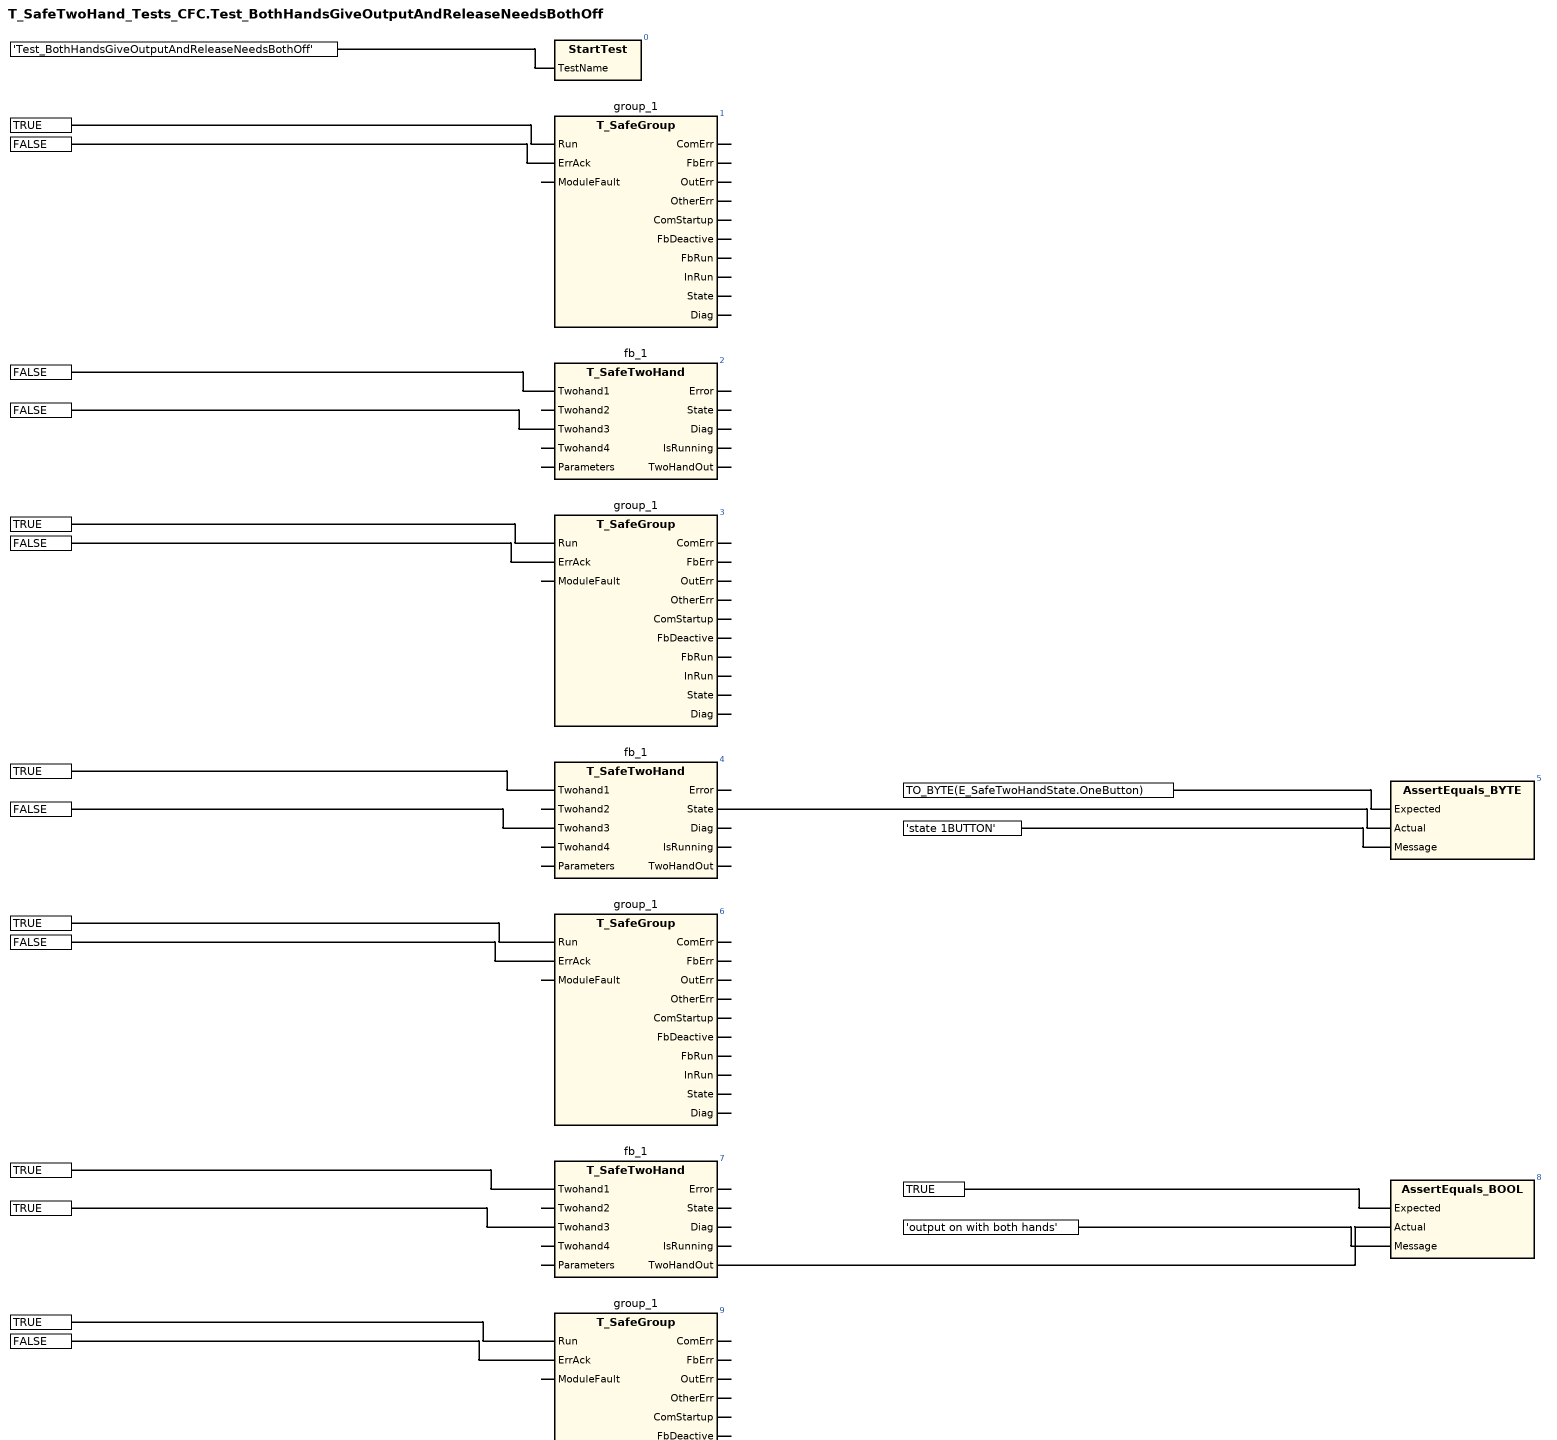
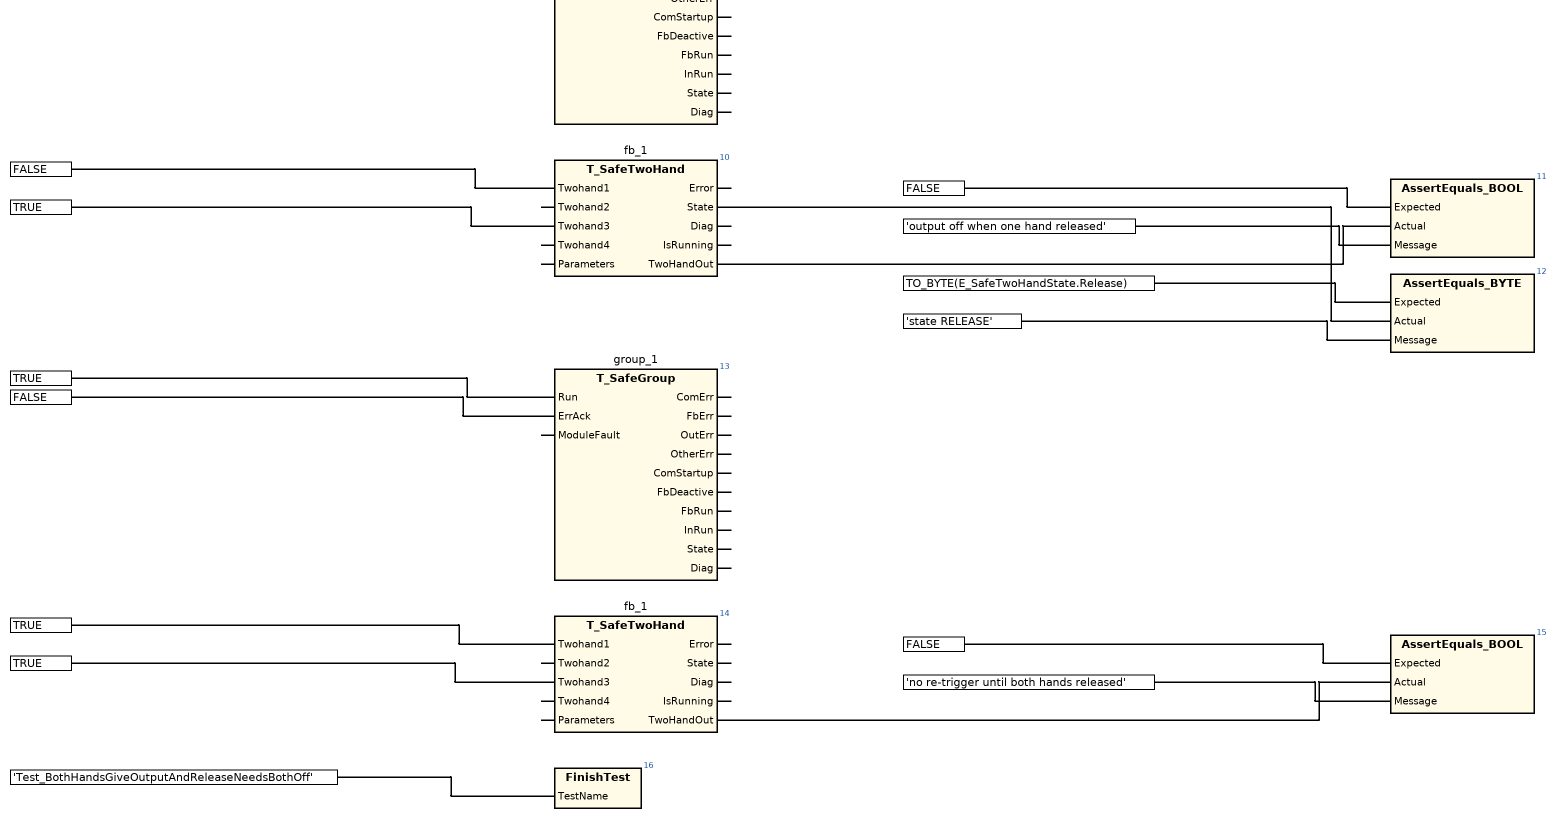
StartTest(TestName := 'Test_BothHandsGiveOutputAndReleaseNeedsBothOff');
group_1(Run := TRUE, ErrAck := FALSE); // T_SafeGroup
fb_1(Twohand1 := FALSE, Twohand3 := FALSE); // T_SafeTwoHand
group_1(Run := TRUE, ErrAck := FALSE); // T_SafeGroup
fb_1(Twohand1 := TRUE, Twohand3 := FALSE); // T_SafeTwoHand
AssertEquals_BYTE(Expected := TO_BYTE(E_SafeTwoHandState.OneButton), Actual := fb_1.State, Message := 'state 1BUTTON');
group_1(Run := TRUE, ErrAck := FALSE); // T_SafeGroup
fb_1(Twohand1 := TRUE, Twohand3 := TRUE); // T_SafeTwoHand
AssertEquals_BOOL(Expected := TRUE, Actual := fb_1.TwoHandOut, Message := 'output on with both hands');
group_1(Run := TRUE, ErrAck := FALSE); // T_SafeGroup
fb_1(Twohand1 := FALSE, Twohand3 := TRUE); // T_SafeTwoHand
AssertEquals_BOOL(Expected := FALSE, Actual := fb_1.TwoHandOut, Message := 'output off when one hand released');
AssertEquals_BYTE(Expected := TO_BYTE(E_SafeTwoHandState.Release), Actual := fb_1.State, Message := 'state RELEASE');
group_1(Run := TRUE, ErrAck := FALSE); // T_SafeGroup
fb_1(Twohand1 := TRUE, Twohand3 := TRUE); // T_SafeTwoHand
AssertEquals_BOOL(Expected := FALSE, Actual := fb_1.TwoHandOut, Message := 'no re-trigger until both hands released');
FinishTest(TestName := 'Test_BothHandsGiveOutputAndReleaseNeedsBothOff');
END_METHOD

METHOD PRIVATE Test_HandDiscrepancyTimeout
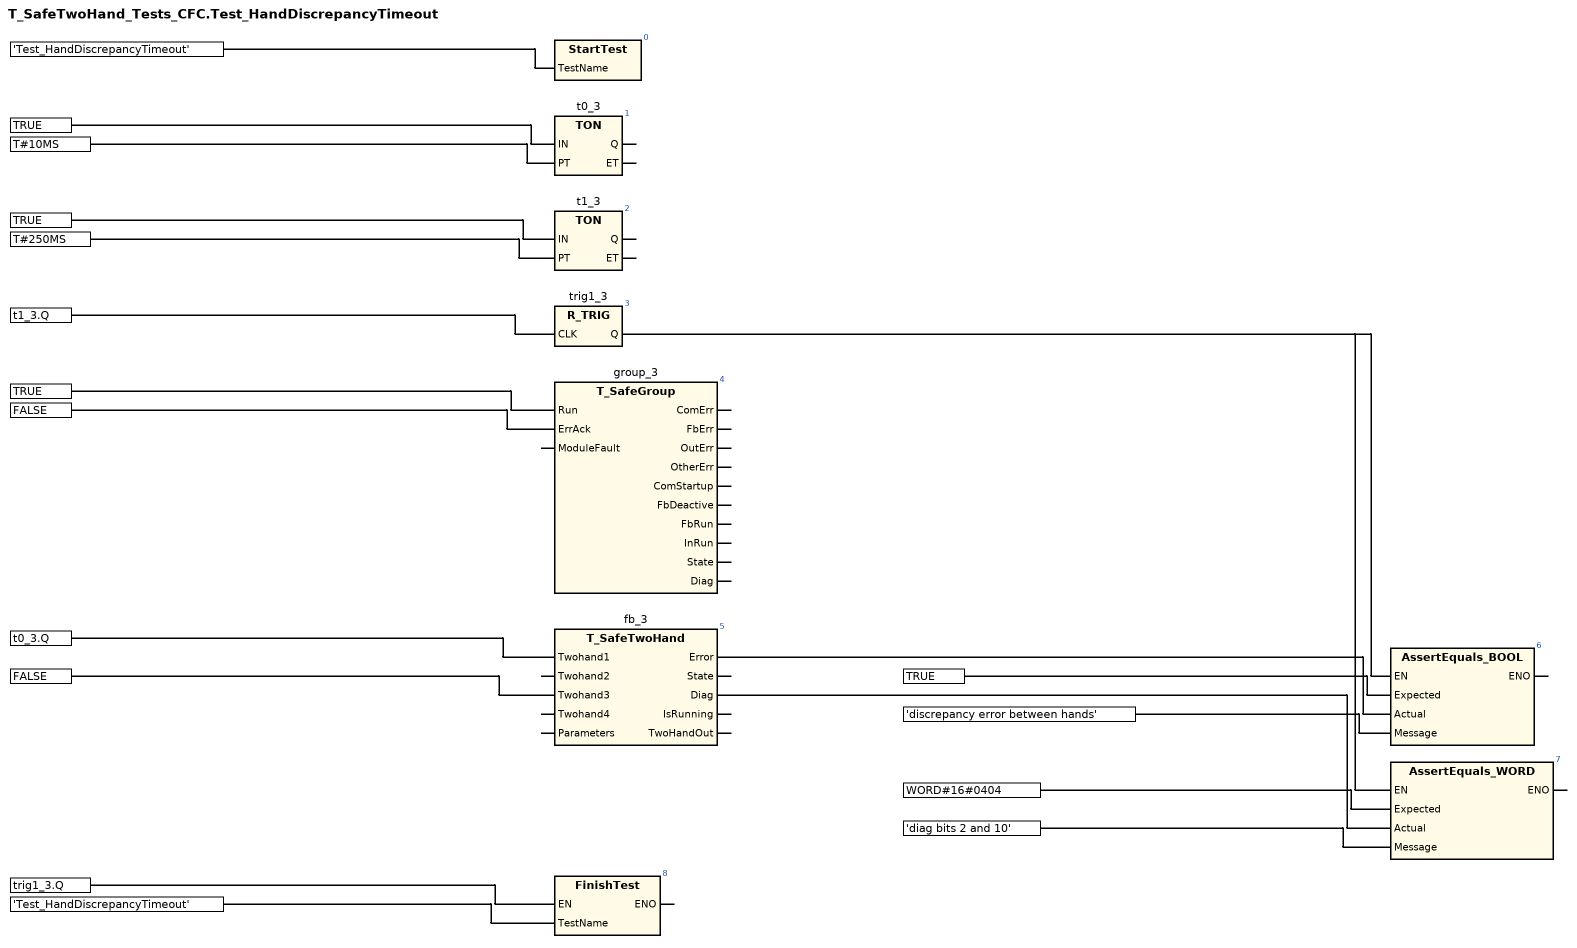
StartTest(TestName := 'Test_HandDiscrepancyTimeout');
t0_3(IN := TRUE, PT := T#10MS); // TON
t1_3(IN := TRUE, PT := T#250MS); // TON
trig1_3(CLK := t1_3.Q); // R_TRIG
group_3(Run := TRUE, ErrAck := FALSE); // T_SafeGroup
fb_3(Twohand1 := t0_3.Q, Twohand3 := FALSE); // T_SafeTwoHand
IF trig1_3.Q THEN AssertEquals_BOOL(Expected := TRUE, Actual := fb_3.Error, Message := 'discrepancy error between hands'); END_IF
IF trig1_3.Q THEN AssertEquals_WORD(Expected := WORD#16#0404, Actual := fb_3.Diag, Message := 'diag bits 2 and 10'); END_IF
IF trig1_3.Q THEN FinishTest(TestName := 'Test_HandDiscrepancyTimeout'); END_IF
END_METHOD

METHOD PRIVATE Test_SecondHandWithoutFirstGivesTwoHandError
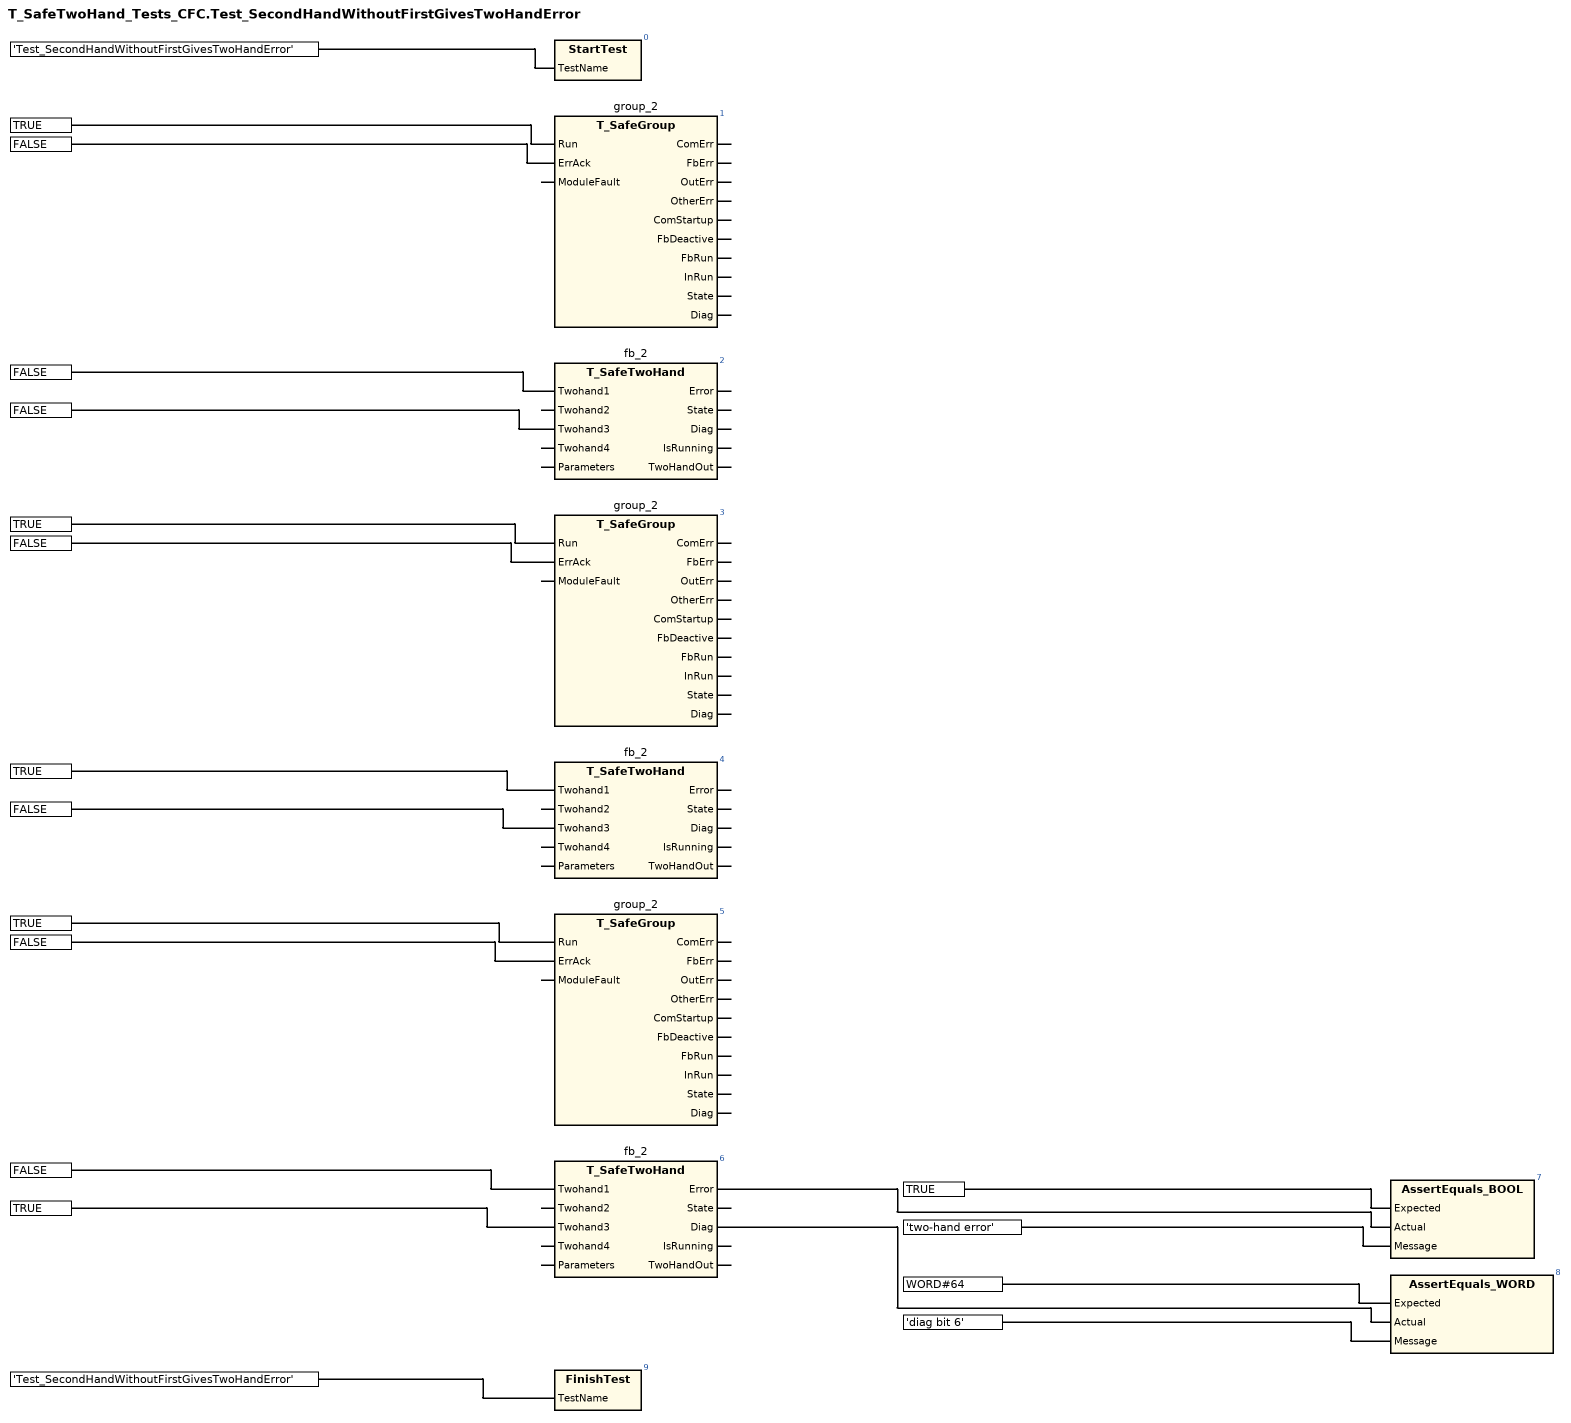
StartTest(TestName := 'Test_SecondHandWithoutFirstGivesTwoHandError');
group_2(Run := TRUE, ErrAck := FALSE); // T_SafeGroup
fb_2(Twohand1 := FALSE, Twohand3 := FALSE); // T_SafeTwoHand
group_2(Run := TRUE, ErrAck := FALSE); // T_SafeGroup
fb_2(Twohand1 := TRUE, Twohand3 := FALSE); // T_SafeTwoHand
group_2(Run := TRUE, ErrAck := FALSE); // T_SafeGroup
fb_2(Twohand1 := FALSE, Twohand3 := TRUE); // T_SafeTwoHand
AssertEquals_BOOL(Expected := TRUE, Actual := fb_2.Error, Message := 'two-hand error');
AssertEquals_WORD(Expected := WORD#64, Actual := fb_2.Diag, Message := 'diag bit 6');
FinishTest(TestName := 'Test_SecondHandWithoutFirstGivesTwoHandError');
END_METHOD

END_FUNCTION_BLOCK

// Tests/T_SafeMuting_Tests_CFC
    // CFC twin of T_SafeMuting_Tests: the same tests drawn as CFC diagrams, the way a TwinSAFE project is authored.
    FUNCTION_BLOCK T_SafeMuting_Tests_CFC EXTENDS T_SafeCfcTestSuite
    VAR
    // Test_OssdBlockedWithoutMutingGivesSafe
    group_1 : T_SafeGroup;
    fb_1 : T_SafeMuting(group := group_1);
    // Test_SequentialMutingKeepsOutputOn
    group_2 : T_SafeGroup;
    fb_2 : T_SafeMuting(group := group_2) := (Parameters := (SequentialInputs := TRUE));
    // Test_SequenceViolationGivesError
    group_3 : T_SafeGroup;
    fb_3 : T_SafeMuting(group := group_3) := (Parameters := (SequentialInputs := TRUE));
    // Test_TwoSensorParallelSequence
    group_4 : T_SafeGroup;
    fb_4 : T_SafeMuting(group := group_4);
END_VAR

Test_OssdBlockedWithoutMutingGivesSafe();
Test_SequentialMutingKeepsOutputOn();
Test_SequenceViolationGivesError();
Test_TwoSensorParallelSequence();

METHOD PRIVATE Test_OssdBlockedWithoutMutingGivesSafe
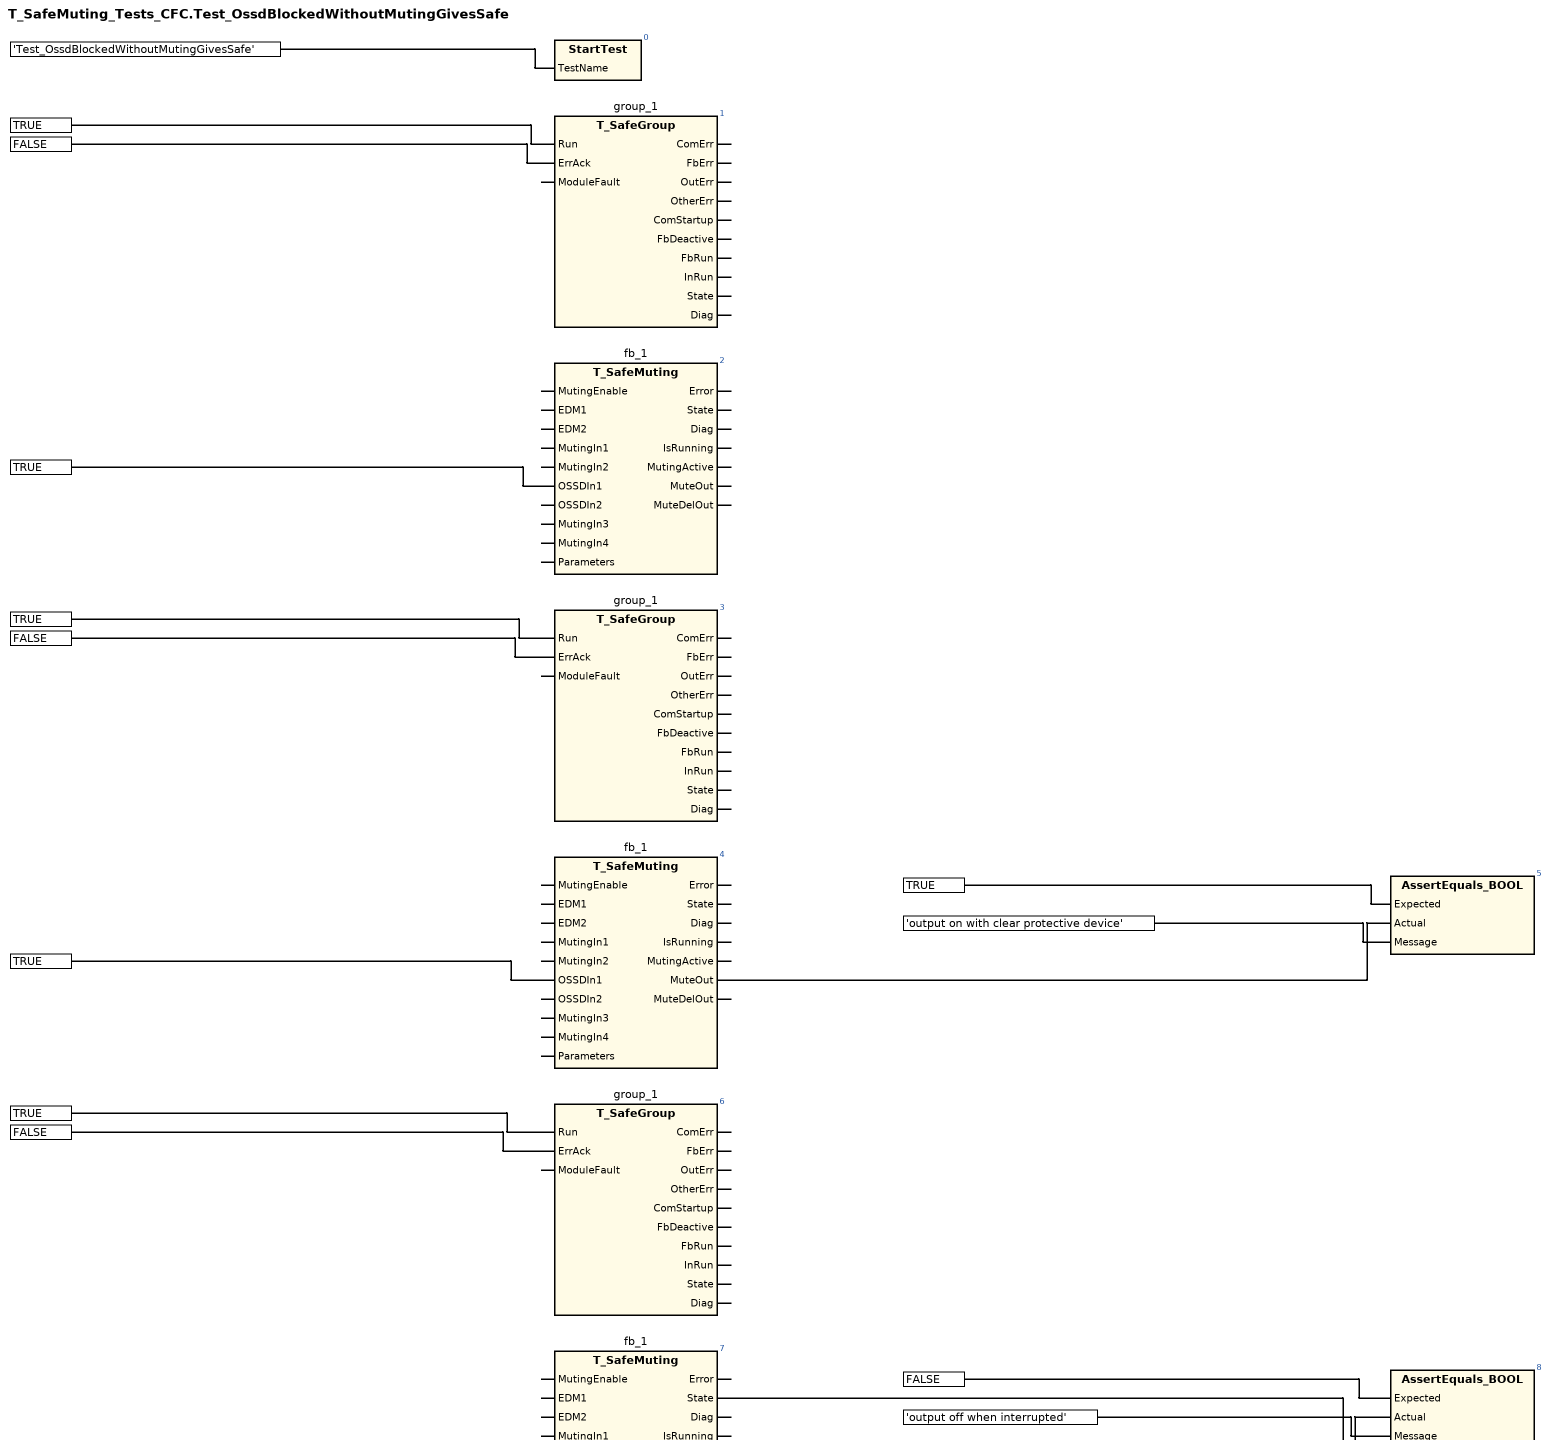
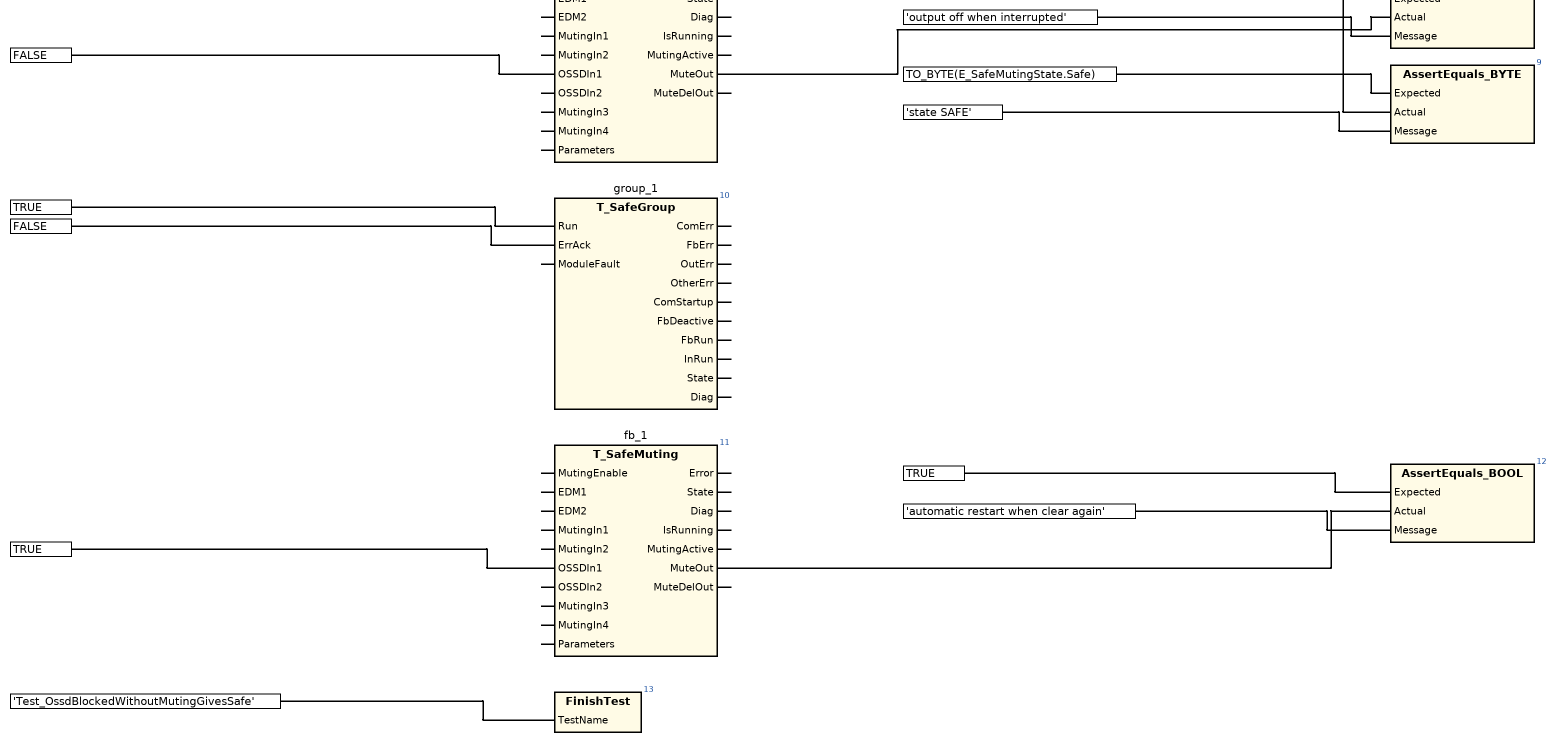
StartTest(TestName := 'Test_OssdBlockedWithoutMutingGivesSafe');
group_1(Run := TRUE, ErrAck := FALSE); // T_SafeGroup
fb_1(OSSDIn1 := TRUE); // T_SafeMuting
group_1(Run := TRUE, ErrAck := FALSE); // T_SafeGroup
fb_1(OSSDIn1 := TRUE); // T_SafeMuting
AssertEquals_BOOL(Expected := TRUE, Actual := fb_1.MuteOut, Message := 'output on with clear protective device');
group_1(Run := TRUE, ErrAck := FALSE); // T_SafeGroup
fb_1(OSSDIn1 := FALSE); // T_SafeMuting
AssertEquals_BOOL(Expected := FALSE, Actual := fb_1.MuteOut, Message := 'output off when interrupted');
AssertEquals_BYTE(Expected := TO_BYTE(E_SafeMutingState.Safe), Actual := fb_1.State, Message := 'state SAFE');
group_1(Run := TRUE, ErrAck := FALSE); // T_SafeGroup
fb_1(OSSDIn1 := TRUE); // T_SafeMuting
AssertEquals_BOOL(Expected := TRUE, Actual := fb_1.MuteOut, Message := 'automatic restart when clear again');
FinishTest(TestName := 'Test_OssdBlockedWithoutMutingGivesSafe');
END_METHOD

METHOD PRIVATE Test_SequenceViolationGivesError
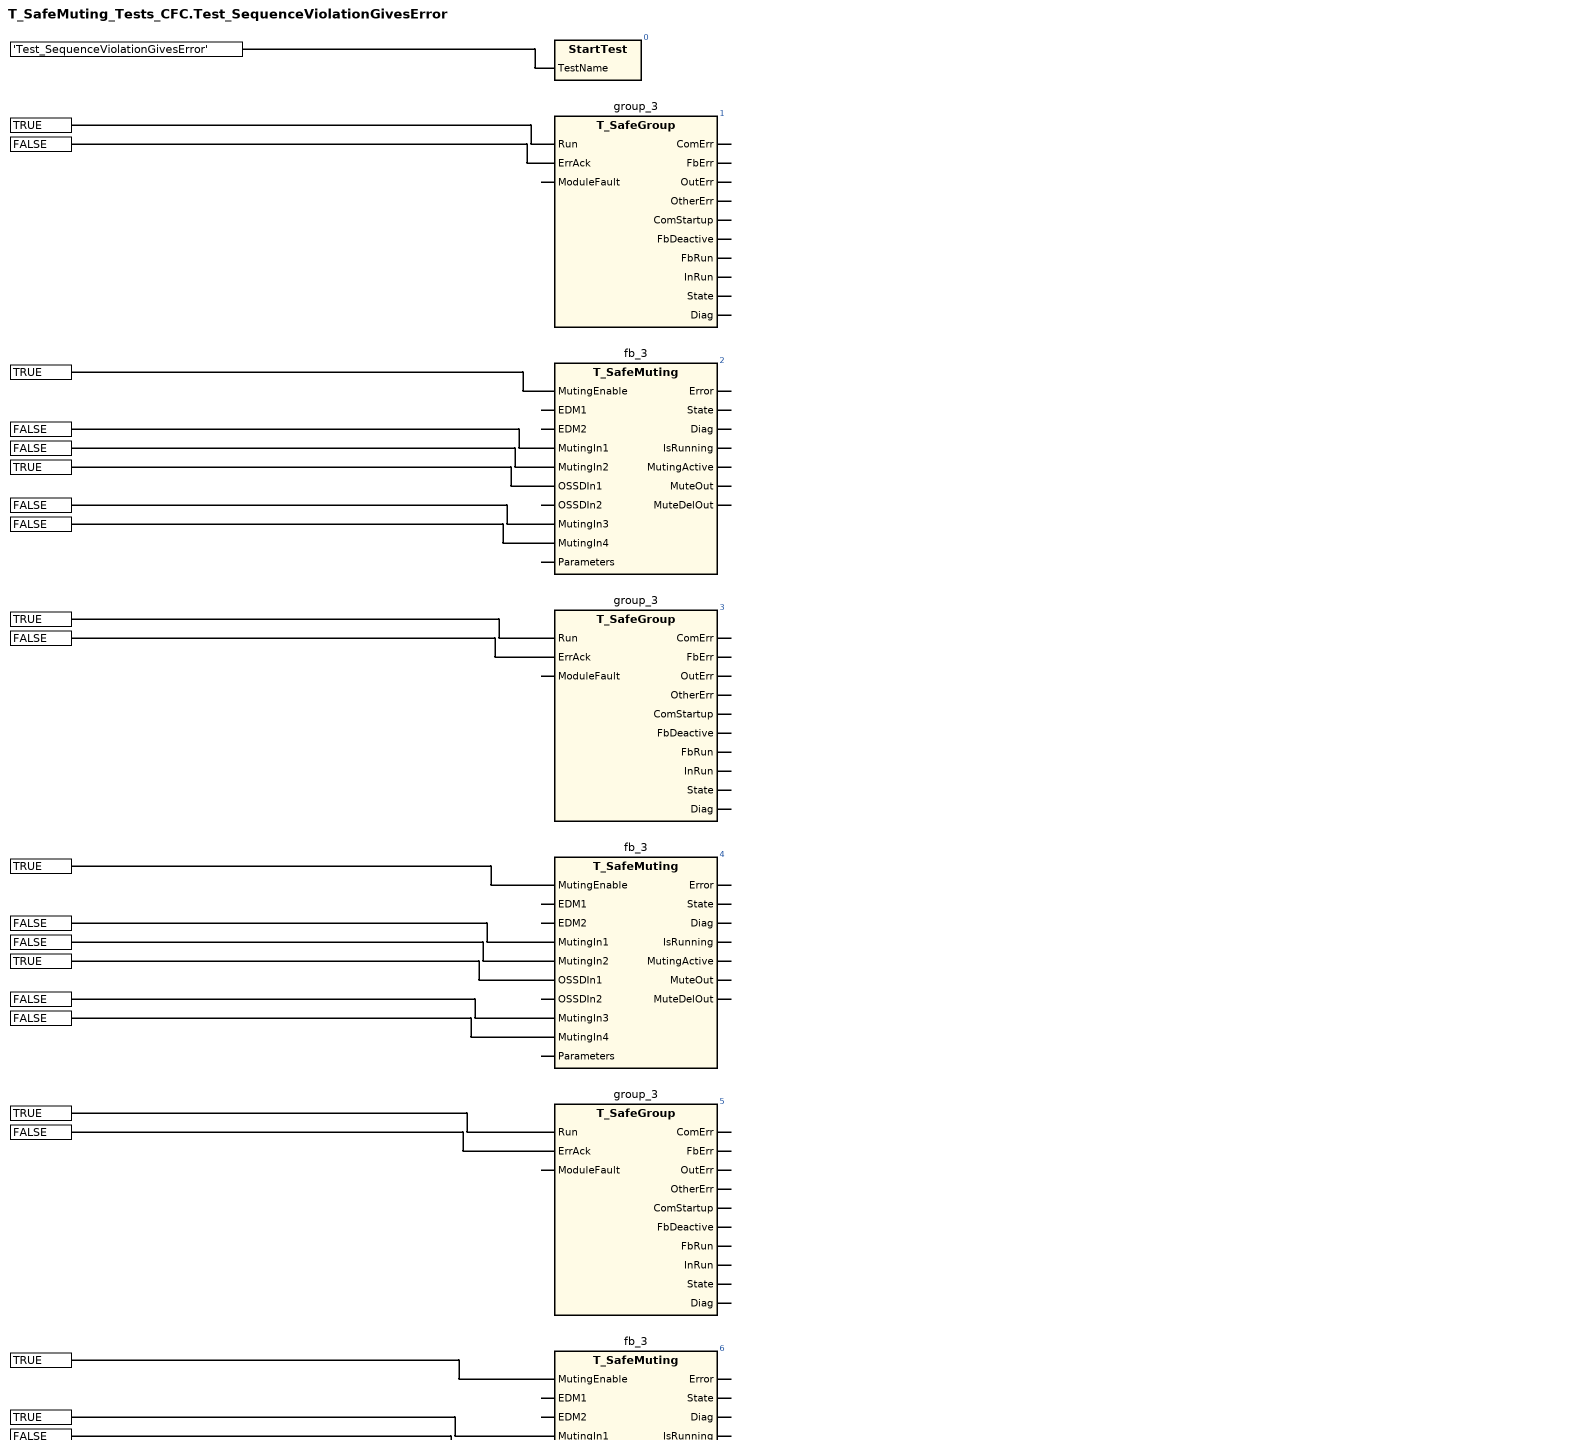
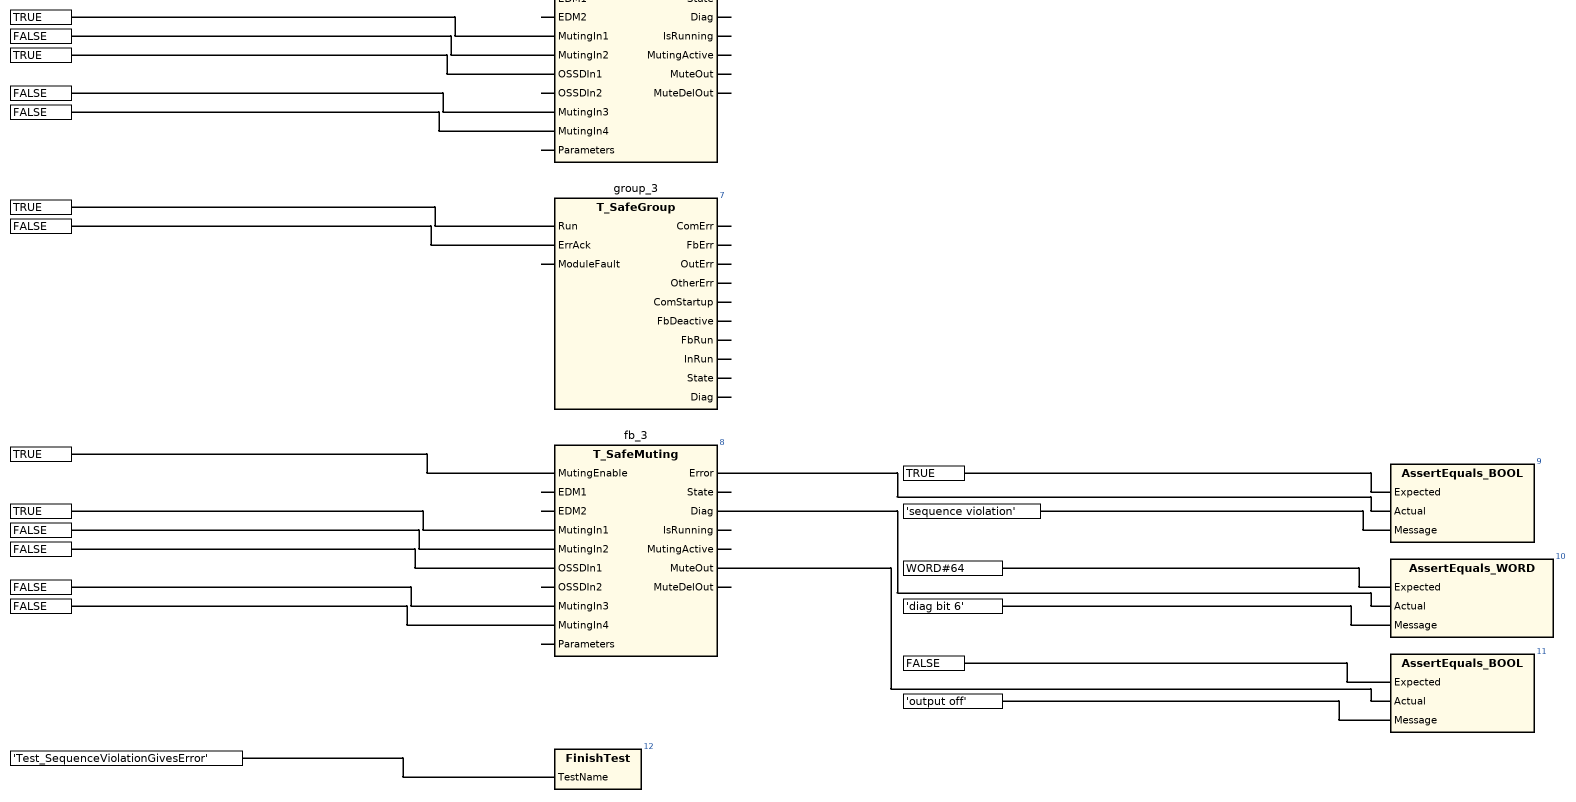
StartTest(TestName := 'Test_SequenceViolationGivesError');
group_3(Run := TRUE, ErrAck := FALSE); // T_SafeGroup
fb_3(
    MutingEnable := TRUE,
    MutingIn1 := FALSE,
    MutingIn2 := FALSE,
    OSSDIn1 := TRUE,
    MutingIn3 := FALSE,
    MutingIn4 := FALSE); // T_SafeMuting
group_3(Run := TRUE, ErrAck := FALSE); // T_SafeGroup
fb_3(
    MutingEnable := TRUE,
    MutingIn1 := FALSE,
    MutingIn2 := FALSE,
    OSSDIn1 := TRUE,
    MutingIn3 := FALSE,
    MutingIn4 := FALSE); // T_SafeMuting
group_3(Run := TRUE, ErrAck := FALSE); // T_SafeGroup
fb_3(
    MutingEnable := TRUE,
    MutingIn1 := TRUE,
    MutingIn2 := FALSE,
    OSSDIn1 := TRUE,
    MutingIn3 := FALSE,
    MutingIn4 := FALSE); // T_SafeMuting
group_3(Run := TRUE, ErrAck := FALSE); // T_SafeGroup
fb_3(
    MutingEnable := TRUE,
    MutingIn1 := TRUE,
    MutingIn2 := FALSE,
    OSSDIn1 := FALSE,
    MutingIn3 := FALSE,
    MutingIn4 := FALSE); // T_SafeMuting
AssertEquals_BOOL(Expected := TRUE, Actual := fb_3.Error, Message := 'sequence violation');
AssertEquals_WORD(Expected := WORD#64, Actual := fb_3.Diag, Message := 'diag bit 6');
AssertEquals_BOOL(Expected := FALSE, Actual := fb_3.MuteOut, Message := 'output off');
FinishTest(TestName := 'Test_SequenceViolationGivesError');
END_METHOD

METHOD PRIVATE Test_SequentialMutingKeepsOutputOn
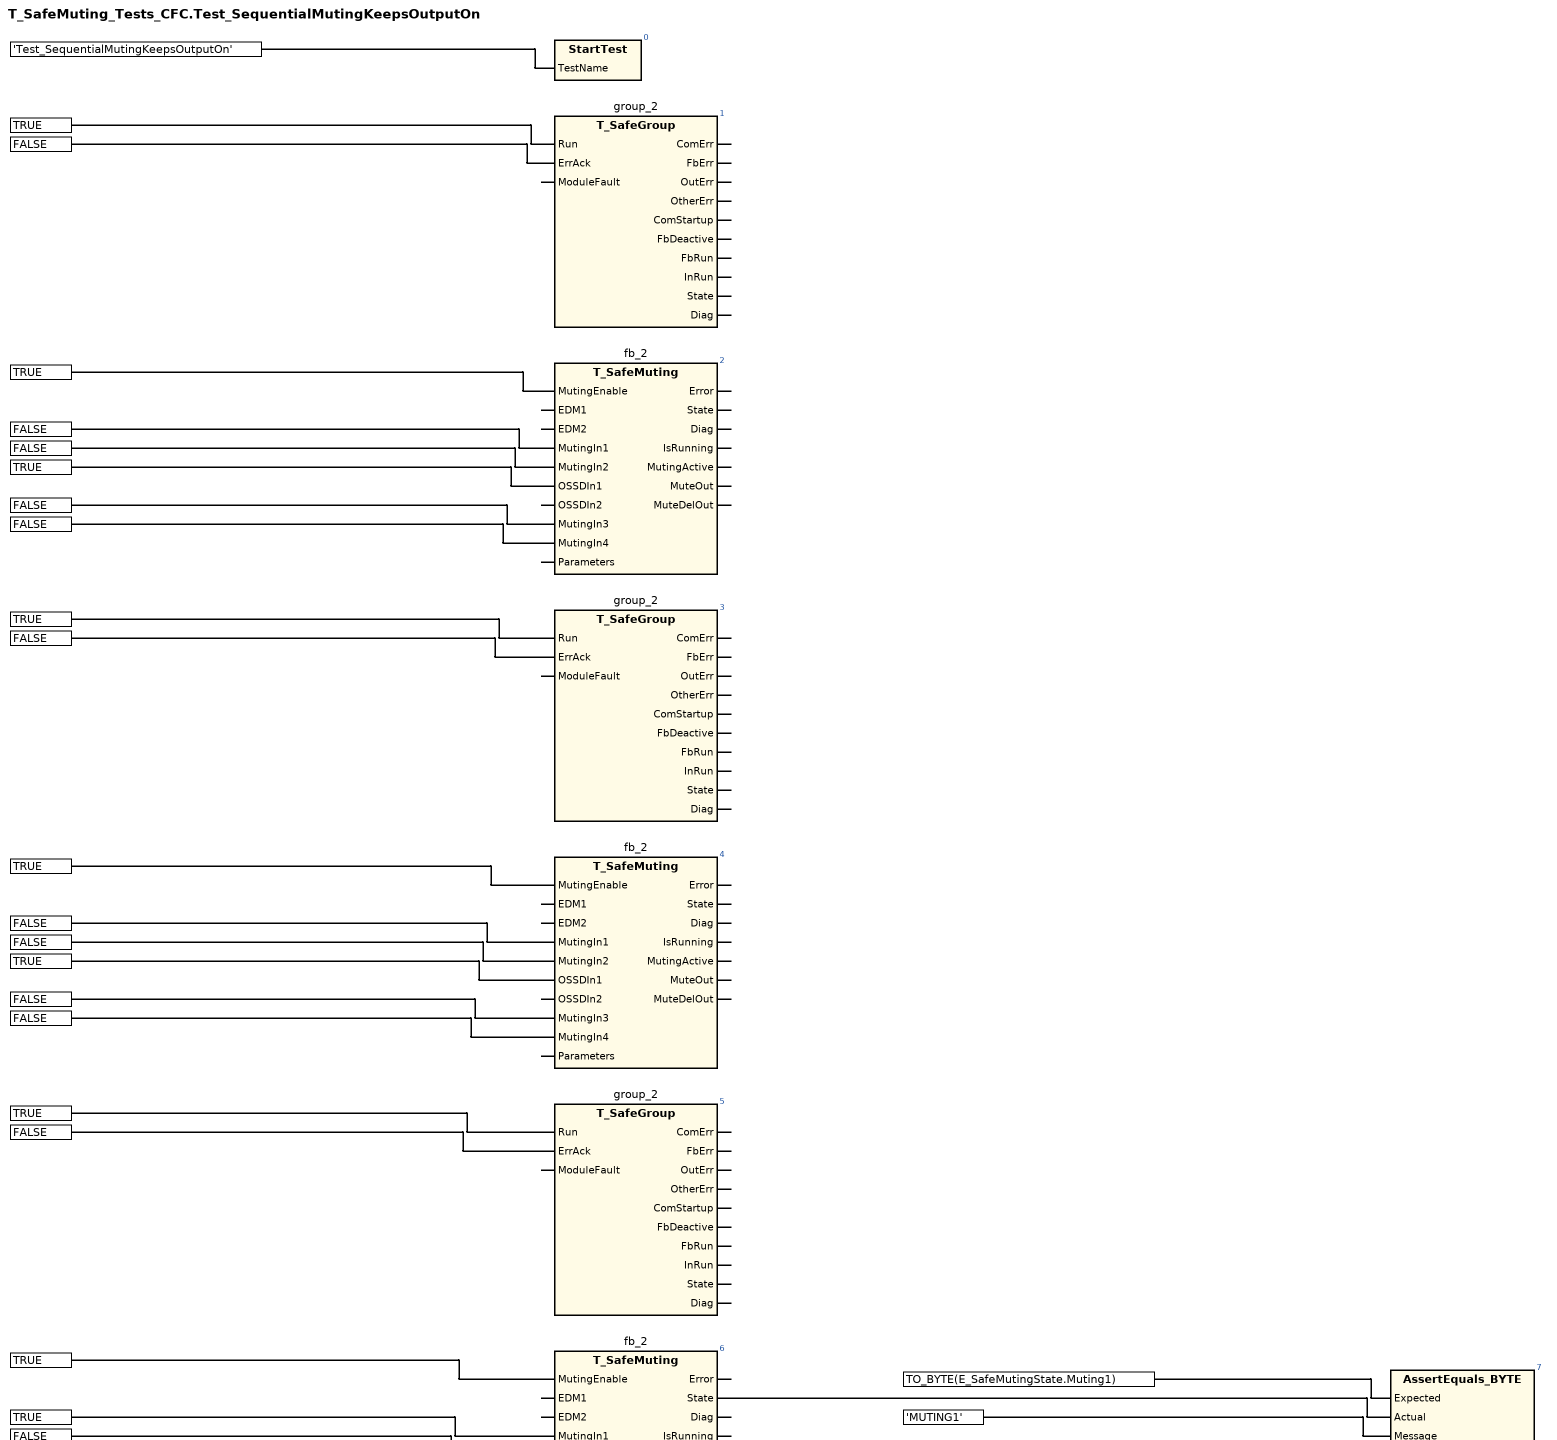
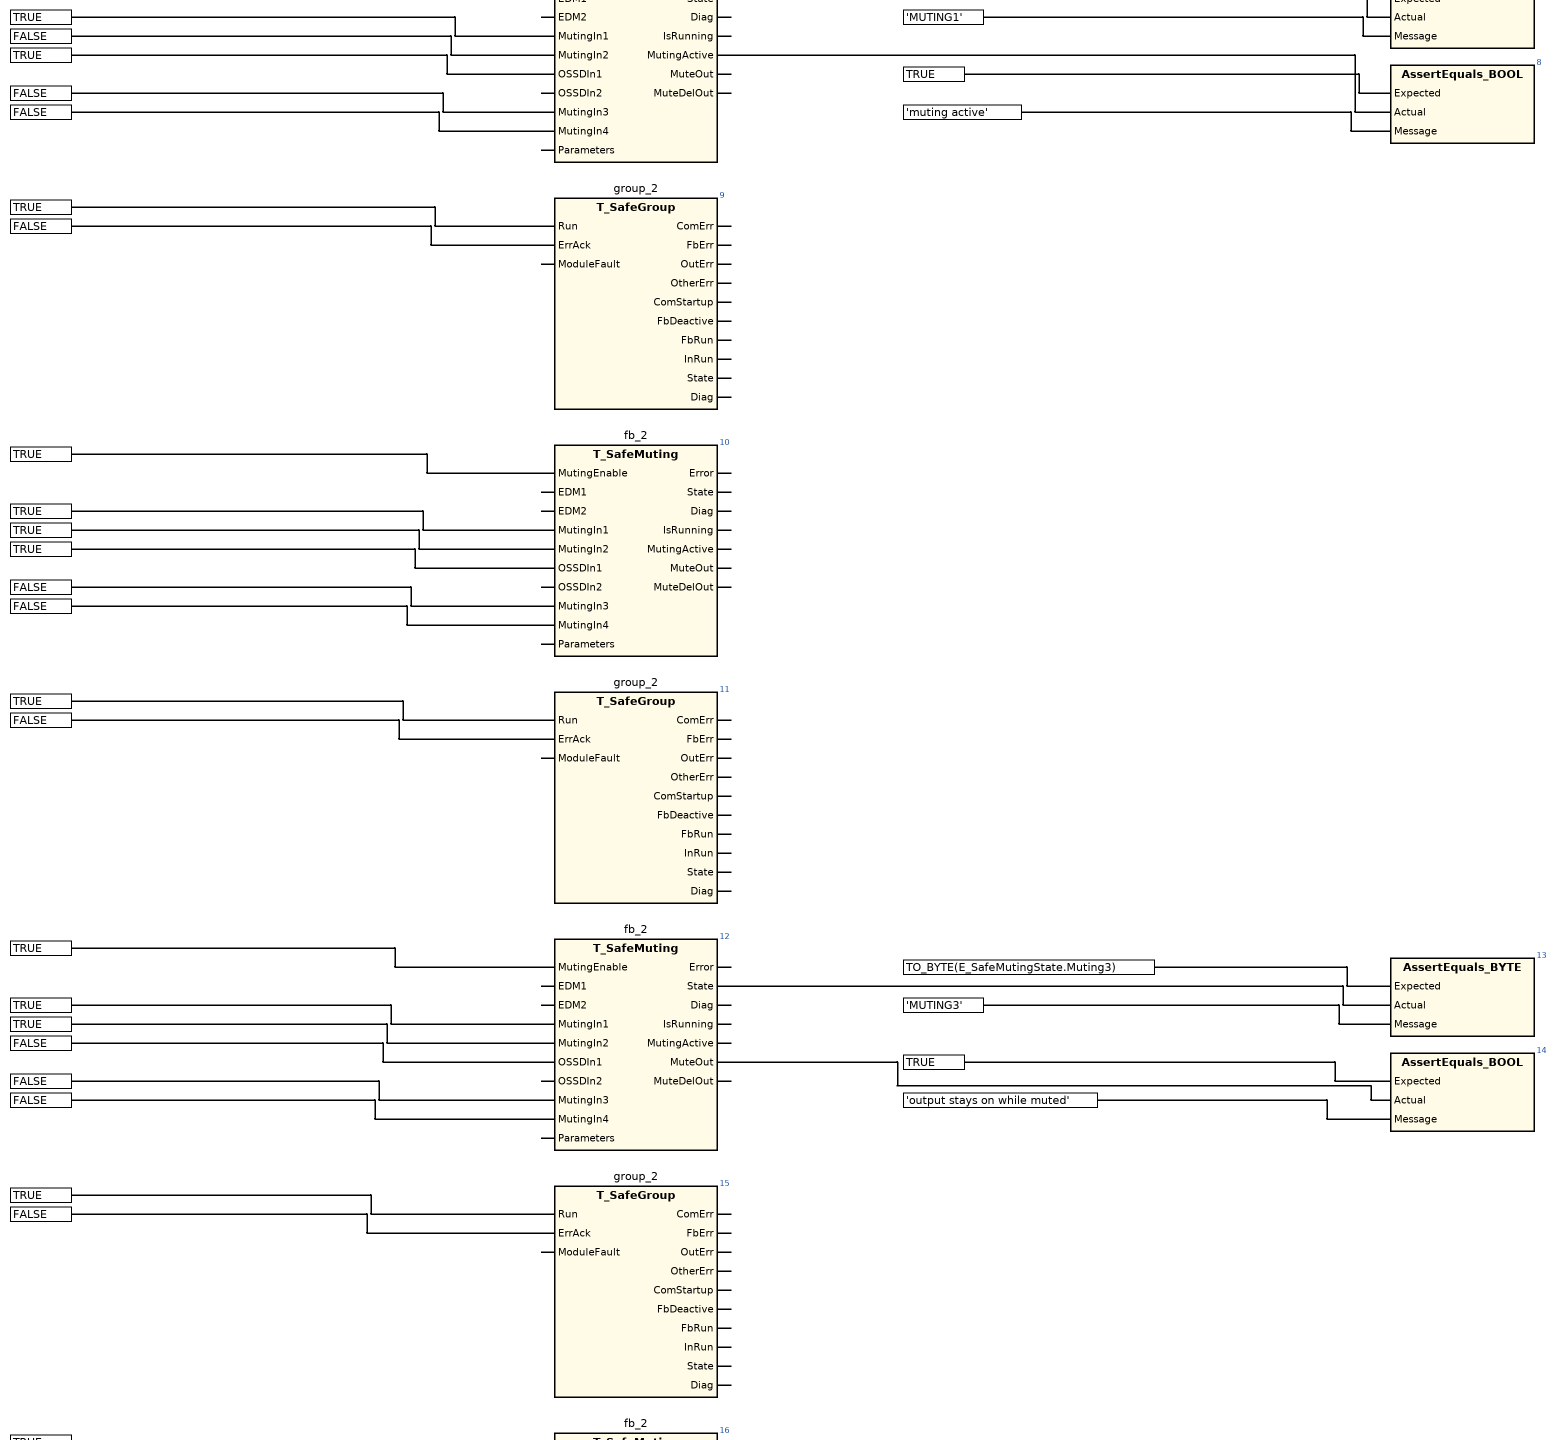
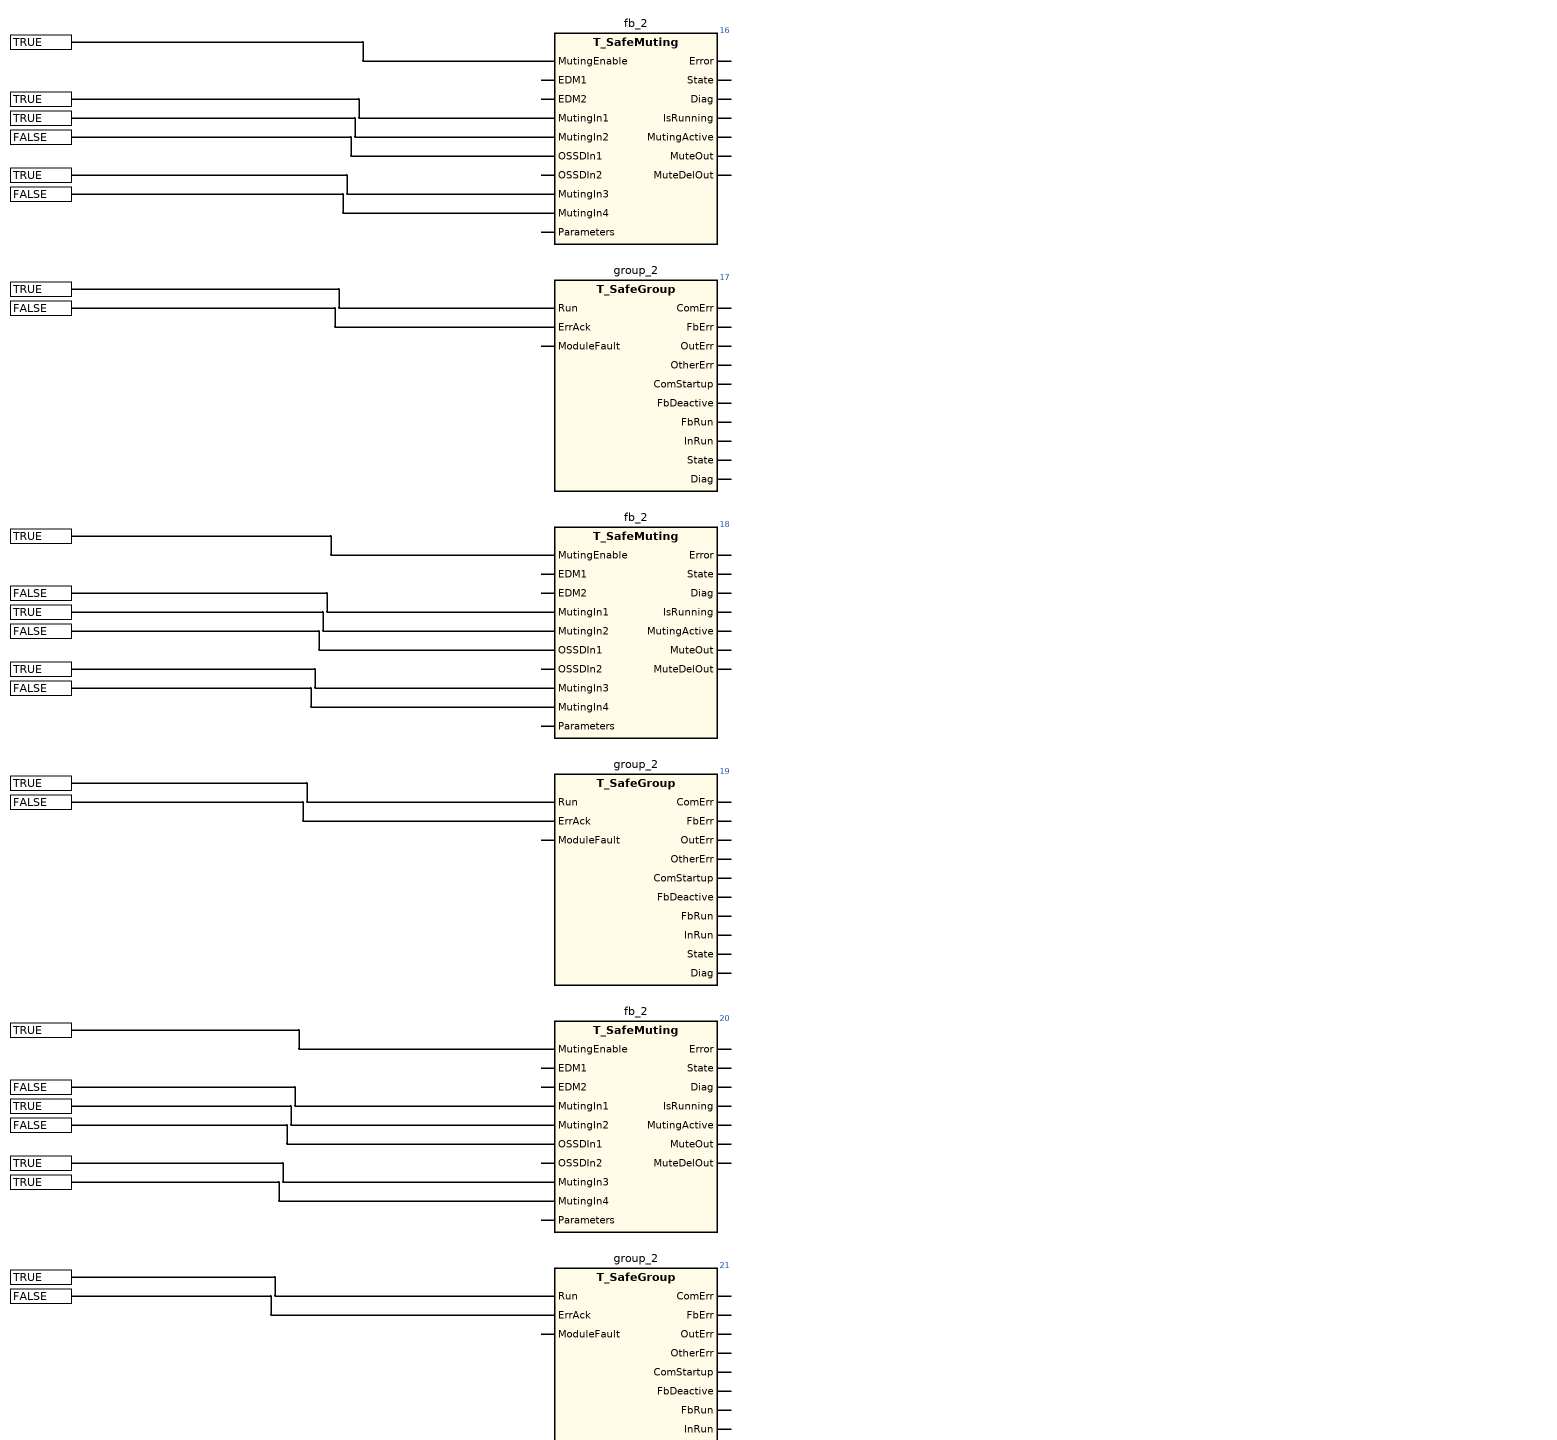
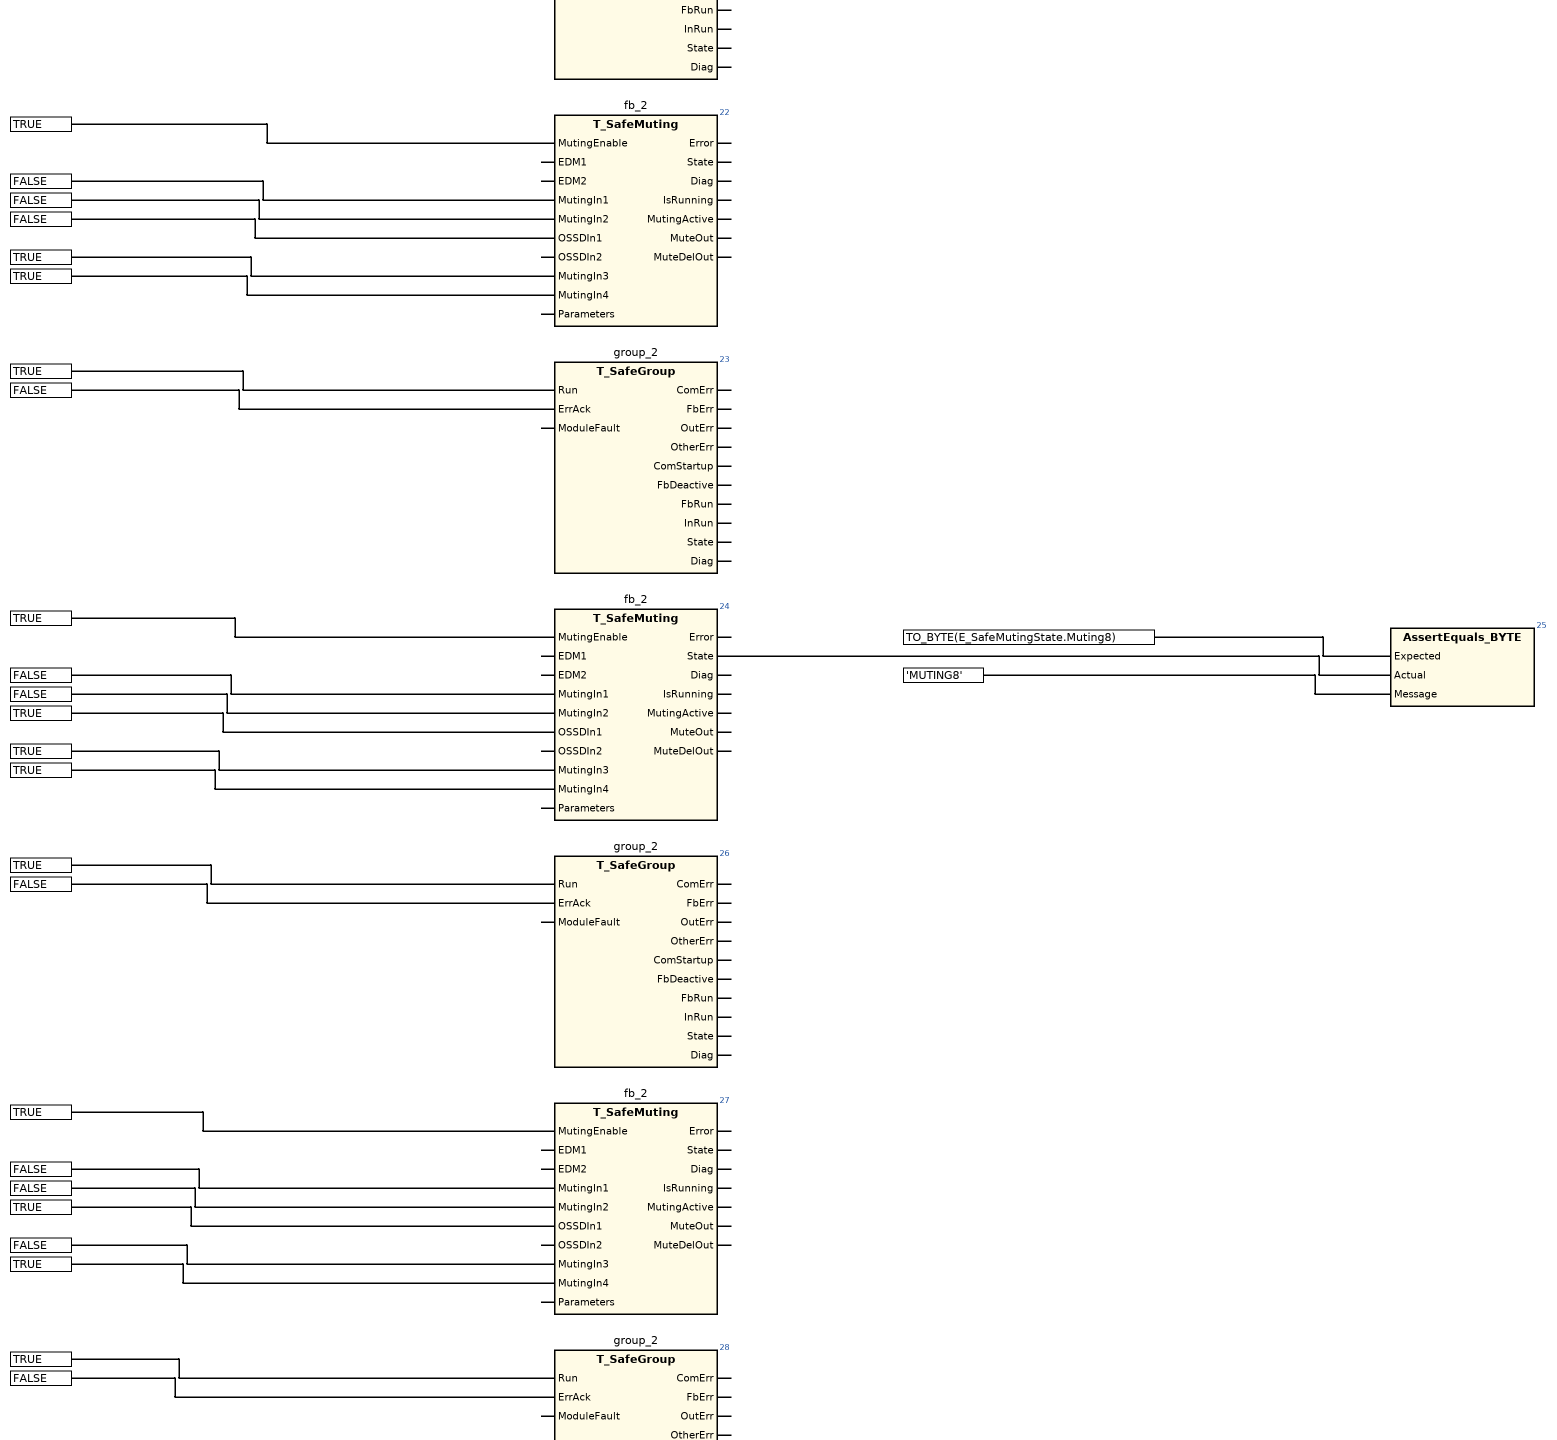
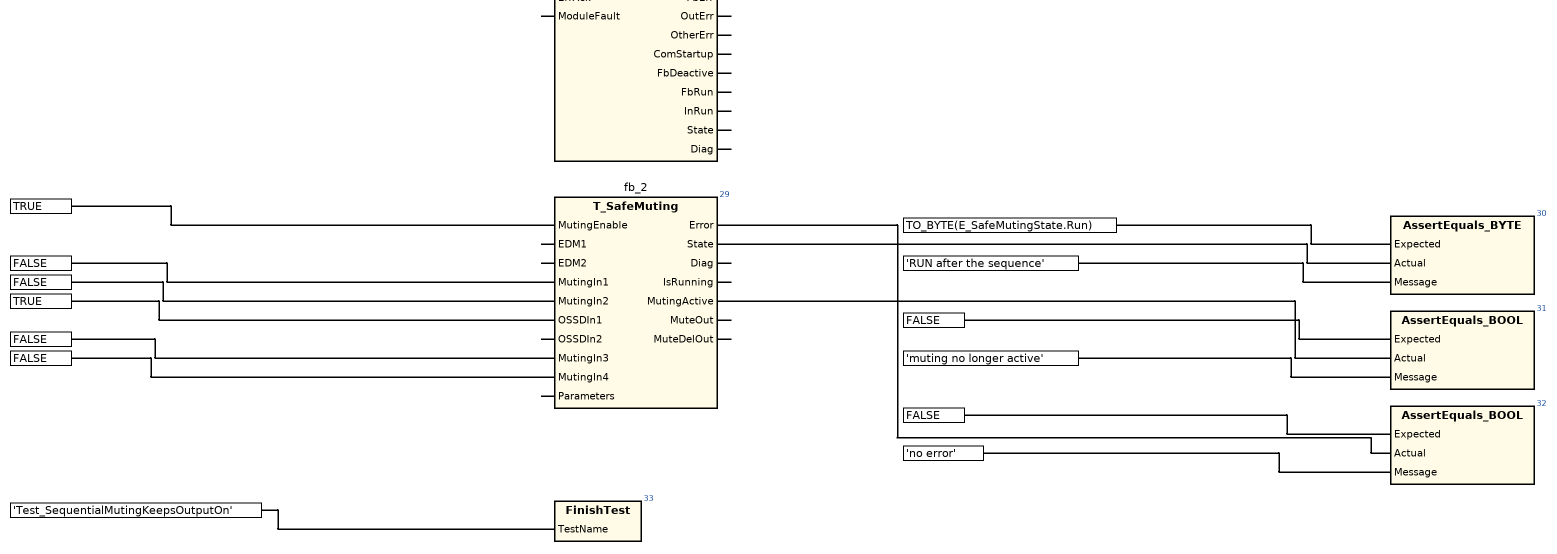
StartTest(TestName := 'Test_SequentialMutingKeepsOutputOn');
group_2(Run := TRUE, ErrAck := FALSE); // T_SafeGroup
fb_2(
    MutingEnable := TRUE,
    MutingIn1 := FALSE,
    MutingIn2 := FALSE,
    OSSDIn1 := TRUE,
    MutingIn3 := FALSE,
    MutingIn4 := FALSE); // T_SafeMuting
group_2(Run := TRUE, ErrAck := FALSE); // T_SafeGroup
fb_2(
    MutingEnable := TRUE,
    MutingIn1 := FALSE,
    MutingIn2 := FALSE,
    OSSDIn1 := TRUE,
    MutingIn3 := FALSE,
    MutingIn4 := FALSE); // T_SafeMuting
group_2(Run := TRUE, ErrAck := FALSE); // T_SafeGroup
fb_2(
    MutingEnable := TRUE,
    MutingIn1 := TRUE,
    MutingIn2 := FALSE,
    OSSDIn1 := TRUE,
    MutingIn3 := FALSE,
    MutingIn4 := FALSE); // T_SafeMuting
AssertEquals_BYTE(Expected := TO_BYTE(E_SafeMutingState.Muting1), Actual := fb_2.State, Message := 'MUTING1');
AssertEquals_BOOL(Expected := TRUE, Actual := fb_2.MutingActive, Message := 'muting active');
group_2(Run := TRUE, ErrAck := FALSE); // T_SafeGroup
fb_2(
    MutingEnable := TRUE,
    MutingIn1 := TRUE,
    MutingIn2 := TRUE,
    OSSDIn1 := TRUE,
    MutingIn3 := FALSE,
    MutingIn4 := FALSE); // T_SafeMuting
group_2(Run := TRUE, ErrAck := FALSE); // T_SafeGroup
fb_2(
    MutingEnable := TRUE,
    MutingIn1 := TRUE,
    MutingIn2 := TRUE,
    OSSDIn1 := FALSE,
    MutingIn3 := FALSE,
    MutingIn4 := FALSE); // T_SafeMuting
AssertEquals_BYTE(Expected := TO_BYTE(E_SafeMutingState.Muting3), Actual := fb_2.State, Message := 'MUTING3');
AssertEquals_BOOL(Expected := TRUE, Actual := fb_2.MuteOut, Message := 'output stays on while muted');
group_2(Run := TRUE, ErrAck := FALSE); // T_SafeGroup
fb_2(
    MutingEnable := TRUE,
    MutingIn1 := TRUE,
    MutingIn2 := TRUE,
    OSSDIn1 := FALSE,
    MutingIn3 := TRUE,
    MutingIn4 := FALSE); // T_SafeMuting
group_2(Run := TRUE, ErrAck := FALSE); // T_SafeGroup
fb_2(
    MutingEnable := TRUE,
    MutingIn1 := FALSE,
    MutingIn2 := TRUE,
    OSSDIn1 := FALSE,
    MutingIn3 := TRUE,
    MutingIn4 := FALSE); // T_SafeMuting
group_2(Run := TRUE, ErrAck := FALSE); // T_SafeGroup
fb_2(
    MutingEnable := TRUE,
    MutingIn1 := FALSE,
    MutingIn2 := TRUE,
    OSSDIn1 := FALSE,
    MutingIn3 := TRUE,
    MutingIn4 := TRUE); // T_SafeMuting
group_2(Run := TRUE, ErrAck := FALSE); // T_SafeGroup
fb_2(
    MutingEnable := TRUE,
    MutingIn1 := FALSE,
    MutingIn2 := FALSE,
    OSSDIn1 := FALSE,
    MutingIn3 := TRUE,
    MutingIn4 := TRUE); // T_SafeMuting
group_2(Run := TRUE, ErrAck := FALSE); // T_SafeGroup
fb_2(
    MutingEnable := TRUE,
    MutingIn1 := FALSE,
    MutingIn2 := FALSE,
    OSSDIn1 := TRUE,
    MutingIn3 := TRUE,
    MutingIn4 := TRUE); // T_SafeMuting
AssertEquals_BYTE(Expected := TO_BYTE(E_SafeMutingState.Muting8), Actual := fb_2.State, Message := 'MUTING8');
group_2(Run := TRUE, ErrAck := FALSE); // T_SafeGroup
fb_2(
    MutingEnable := TRUE,
    MutingIn1 := FALSE,
    MutingIn2 := FALSE,
    OSSDIn1 := TRUE,
    MutingIn3 := FALSE,
    MutingIn4 := TRUE); // T_SafeMuting
group_2(Run := TRUE, ErrAck := FALSE); // T_SafeGroup
fb_2(
    MutingEnable := TRUE,
    MutingIn1 := FALSE,
    MutingIn2 := FALSE,
    OSSDIn1 := TRUE,
    MutingIn3 := FALSE,
    MutingIn4 := FALSE); // T_SafeMuting
AssertEquals_BYTE(Expected := TO_BYTE(E_SafeMutingState.Run), Actual := fb_2.State, Message := 'RUN after the sequence');
AssertEquals_BOOL(Expected := FALSE, Actual := fb_2.MutingActive, Message := 'muting no longer active');
AssertEquals_BOOL(Expected := FALSE, Actual := fb_2.Error, Message := 'no error');
FinishTest(TestName := 'Test_SequentialMutingKeepsOutputOn');
END_METHOD

METHOD PRIVATE Test_TwoSensorParallelSequence
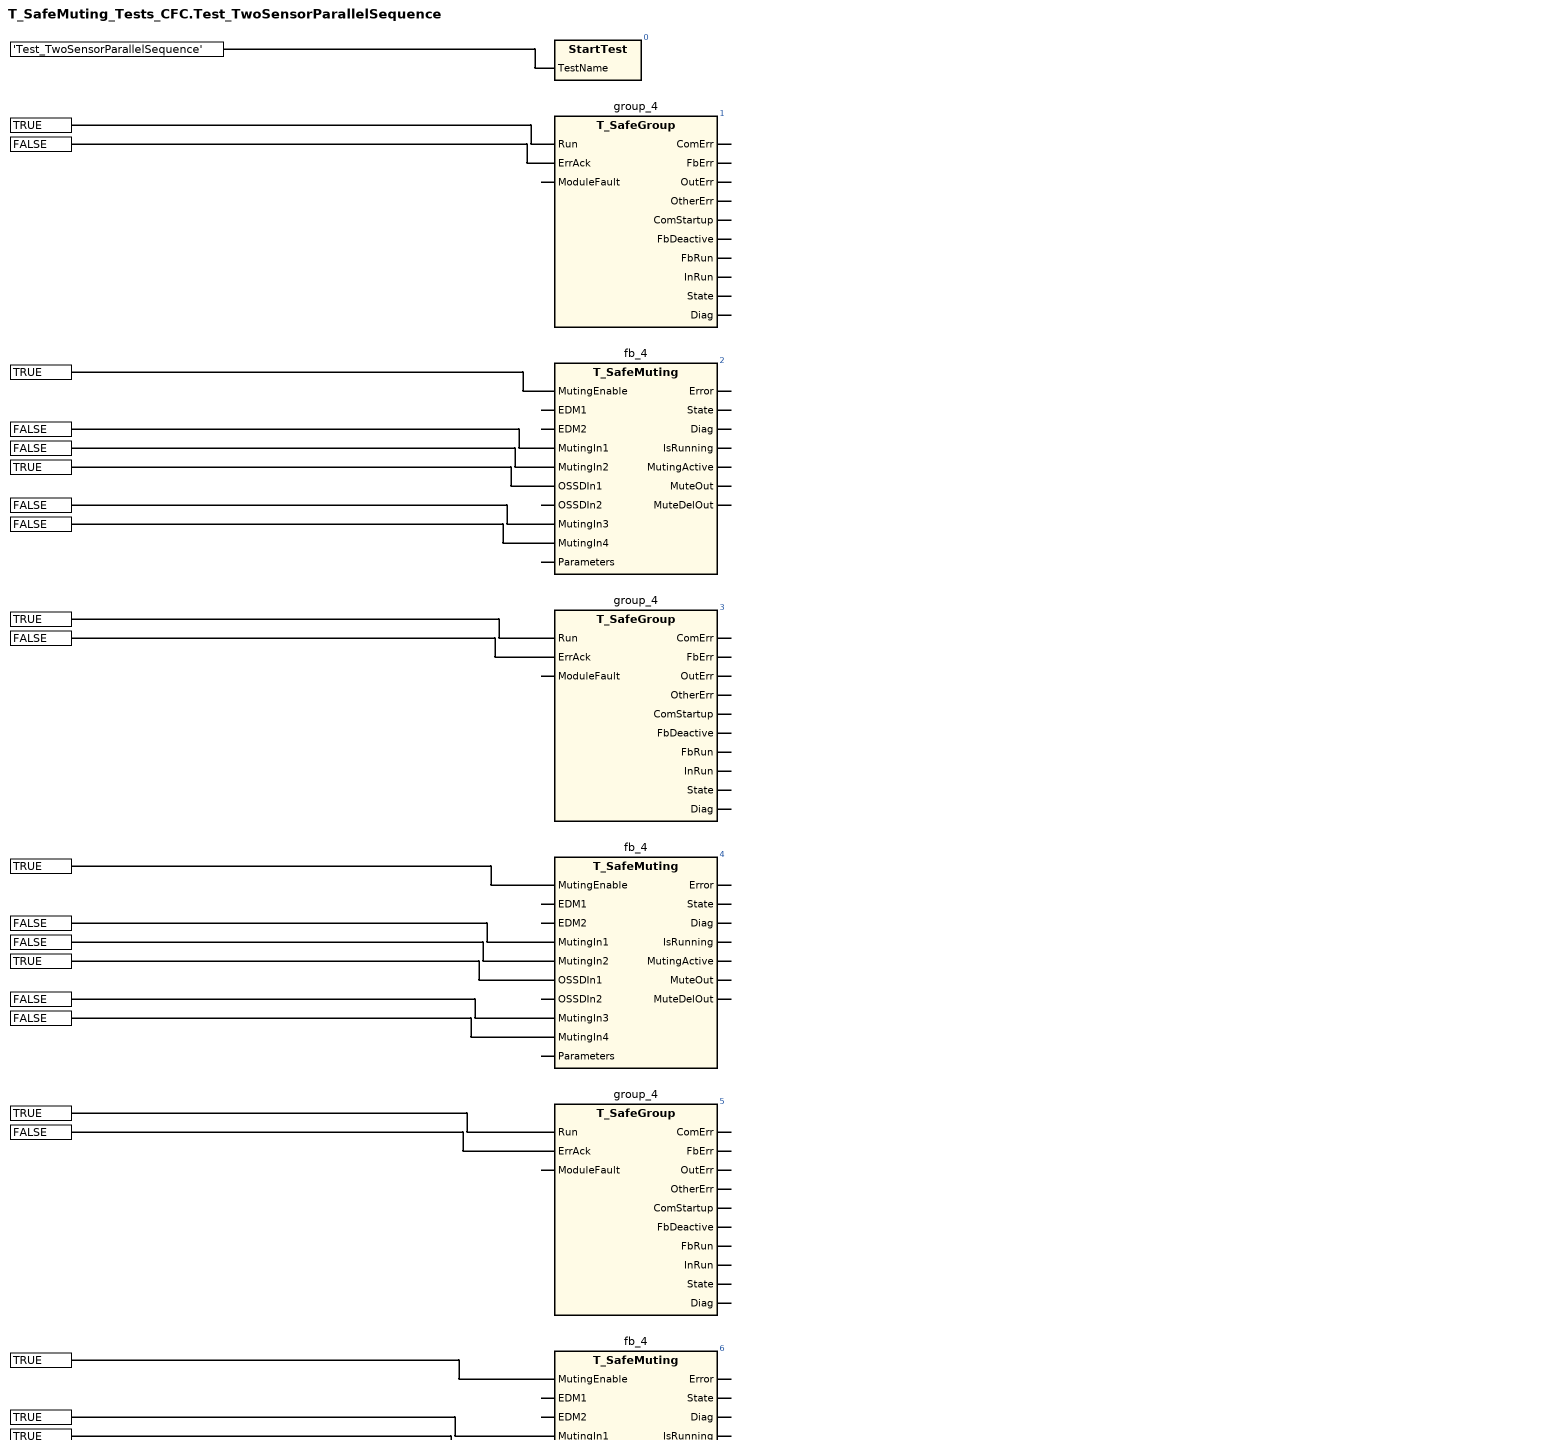
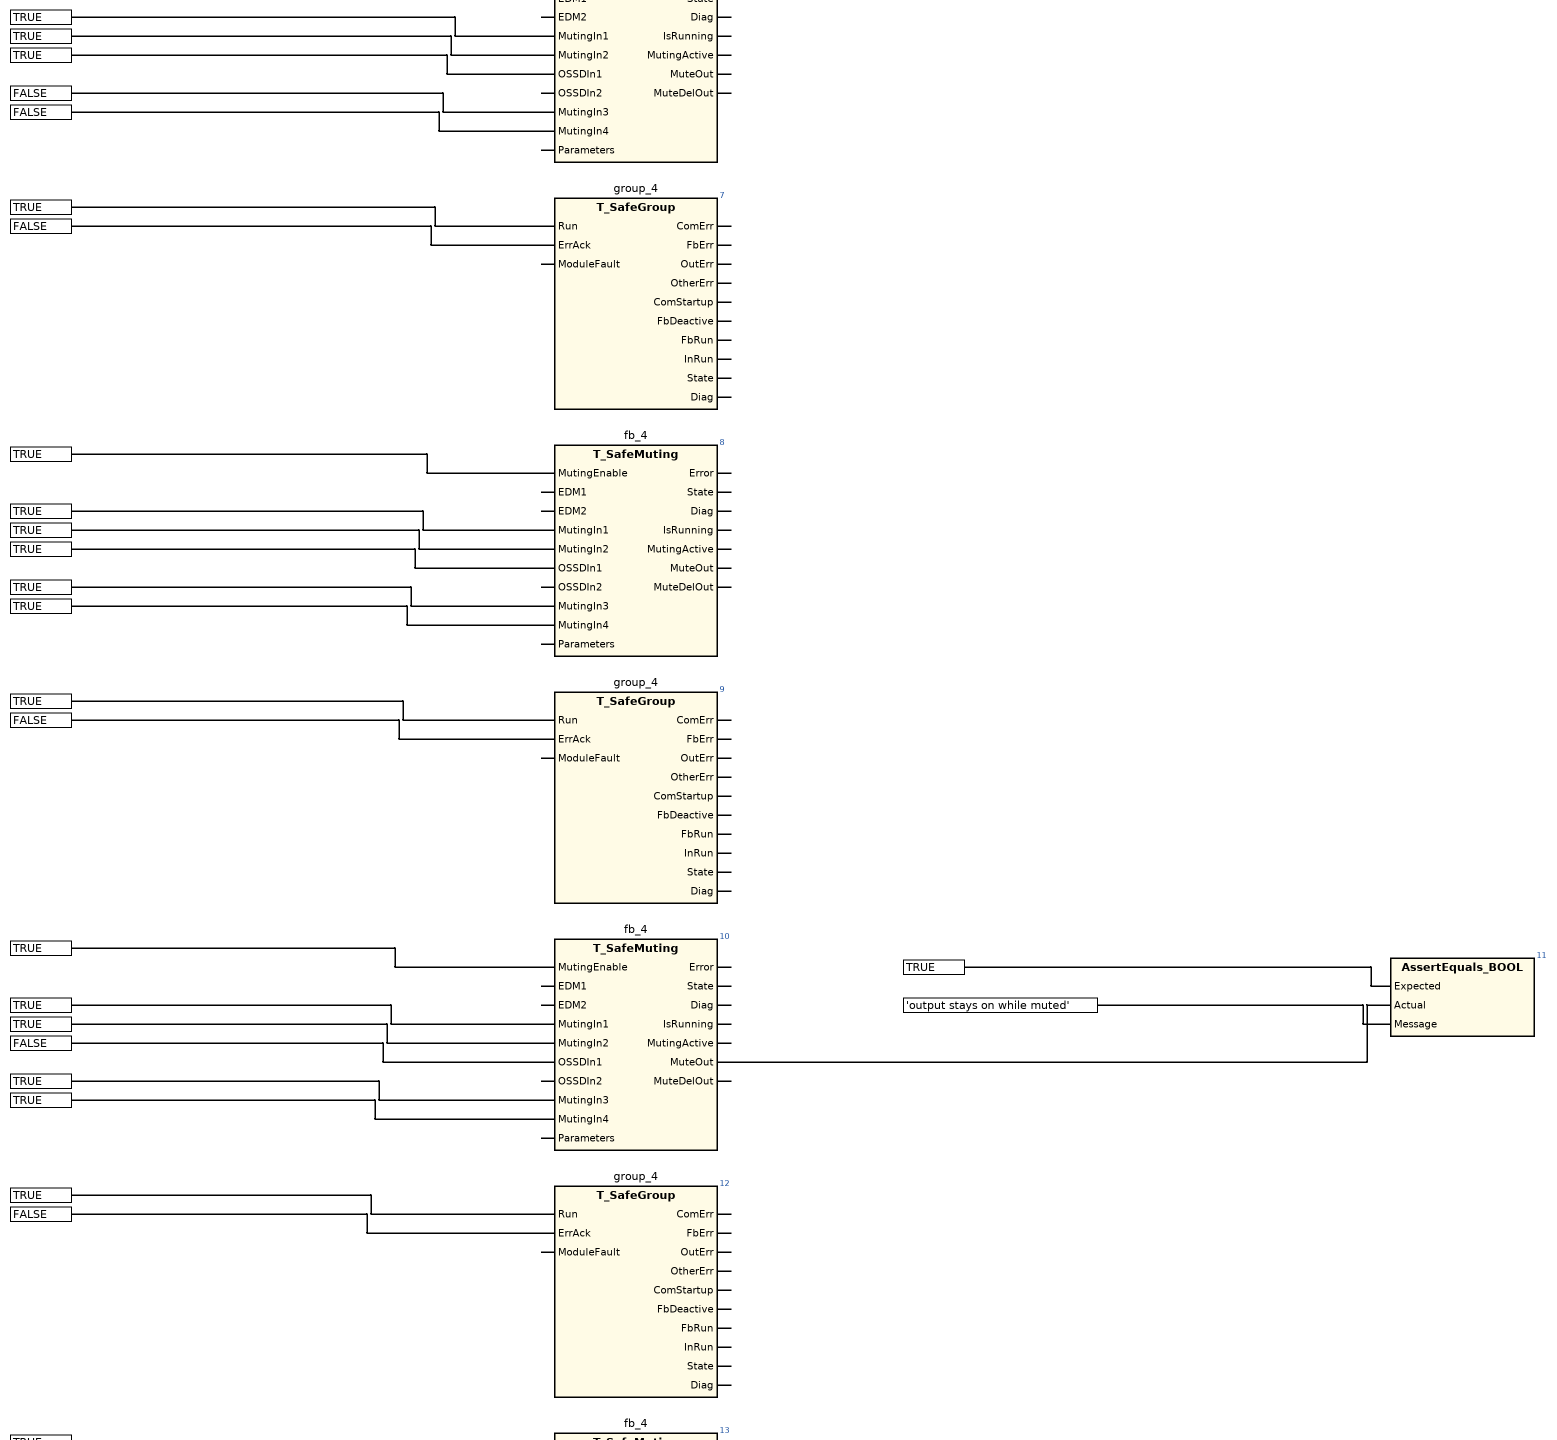
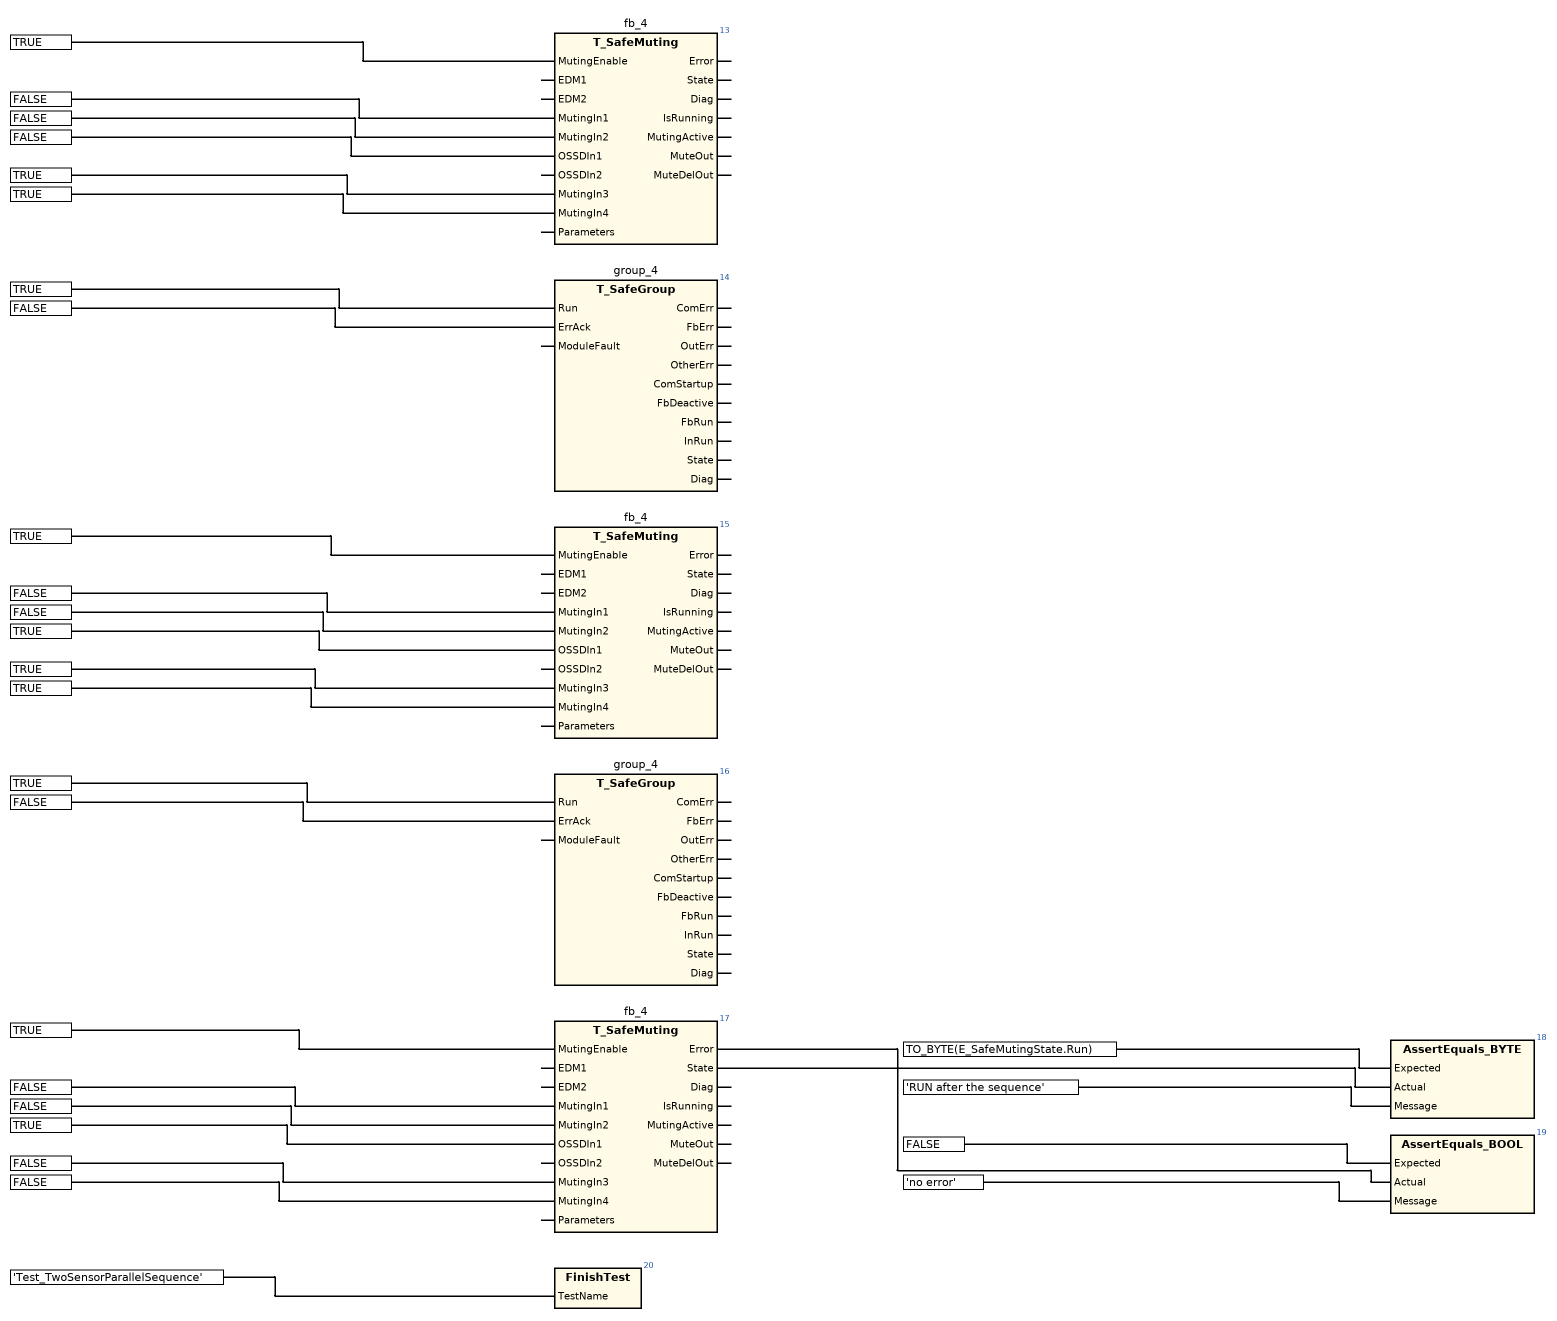
StartTest(TestName := 'Test_TwoSensorParallelSequence');
group_4(Run := TRUE, ErrAck := FALSE); // T_SafeGroup
fb_4(
    MutingEnable := TRUE,
    MutingIn1 := FALSE,
    MutingIn2 := FALSE,
    OSSDIn1 := TRUE,
    MutingIn3 := FALSE,
    MutingIn4 := FALSE); // T_SafeMuting
group_4(Run := TRUE, ErrAck := FALSE); // T_SafeGroup
fb_4(
    MutingEnable := TRUE,
    MutingIn1 := FALSE,
    MutingIn2 := FALSE,
    OSSDIn1 := TRUE,
    MutingIn3 := FALSE,
    MutingIn4 := FALSE); // T_SafeMuting
group_4(Run := TRUE, ErrAck := FALSE); // T_SafeGroup
fb_4(
    MutingEnable := TRUE,
    MutingIn1 := TRUE,
    MutingIn2 := TRUE,
    OSSDIn1 := TRUE,
    MutingIn3 := FALSE,
    MutingIn4 := FALSE); // T_SafeMuting
group_4(Run := TRUE, ErrAck := FALSE); // T_SafeGroup
fb_4(
    MutingEnable := TRUE,
    MutingIn1 := TRUE,
    MutingIn2 := TRUE,
    OSSDIn1 := TRUE,
    MutingIn3 := TRUE,
    MutingIn4 := TRUE); // T_SafeMuting
group_4(Run := TRUE, ErrAck := FALSE); // T_SafeGroup
fb_4(
    MutingEnable := TRUE,
    MutingIn1 := TRUE,
    MutingIn2 := TRUE,
    OSSDIn1 := FALSE,
    MutingIn3 := TRUE,
    MutingIn4 := TRUE); // T_SafeMuting
AssertEquals_BOOL(Expected := TRUE, Actual := fb_4.MuteOut, Message := 'output stays on while muted');
group_4(Run := TRUE, ErrAck := FALSE); // T_SafeGroup
fb_4(
    MutingEnable := TRUE,
    MutingIn1 := FALSE,
    MutingIn2 := FALSE,
    OSSDIn1 := FALSE,
    MutingIn3 := TRUE,
    MutingIn4 := TRUE); // T_SafeMuting
group_4(Run := TRUE, ErrAck := FALSE); // T_SafeGroup
fb_4(
    MutingEnable := TRUE,
    MutingIn1 := FALSE,
    MutingIn2 := FALSE,
    OSSDIn1 := TRUE,
    MutingIn3 := TRUE,
    MutingIn4 := TRUE); // T_SafeMuting
group_4(Run := TRUE, ErrAck := FALSE); // T_SafeGroup
fb_4(
    MutingEnable := TRUE,
    MutingIn1 := FALSE,
    MutingIn2 := FALSE,
    OSSDIn1 := TRUE,
    MutingIn3 := FALSE,
    MutingIn4 := FALSE); // T_SafeMuting
AssertEquals_BYTE(Expected := TO_BYTE(E_SafeMutingState.Run), Actual := fb_4.State, Message := 'RUN after the sequence');
AssertEquals_BOOL(Expected := FALSE, Actual := fb_4.Error, Message := 'no error');
FinishTest(TestName := 'Test_TwoSensorParallelSequence');
END_METHOD

END_FUNCTION_BLOCK

// Tests/T_SafeConnection_Tests_CFC
    // CFC twin of T_SafeConnection_Tests: the same tests drawn as CFC diagrams, the way a TwinSAFE project is authored.
    FUNCTION_BLOCK T_SafeConnection_Tests_CFC EXTENDS T_SafeCfcTestSuite
    VAR
    // Test_StartsUpToDataWhenGroupRuns
    group_1 : T_SafeGroup;
    conn_1 : T_SafeConnection(group := group_1);
    // Test_ComErrorClearedByAcknowledge
    group_2 : T_SafeGroup;
    conn_2 : T_SafeConnection(group := group_2);
END_VAR

Test_StartsUpToDataWhenGroupRuns();
Test_ComErrorClearedByAcknowledge();

METHOD PRIVATE Test_ComErrorClearedByAcknowledge
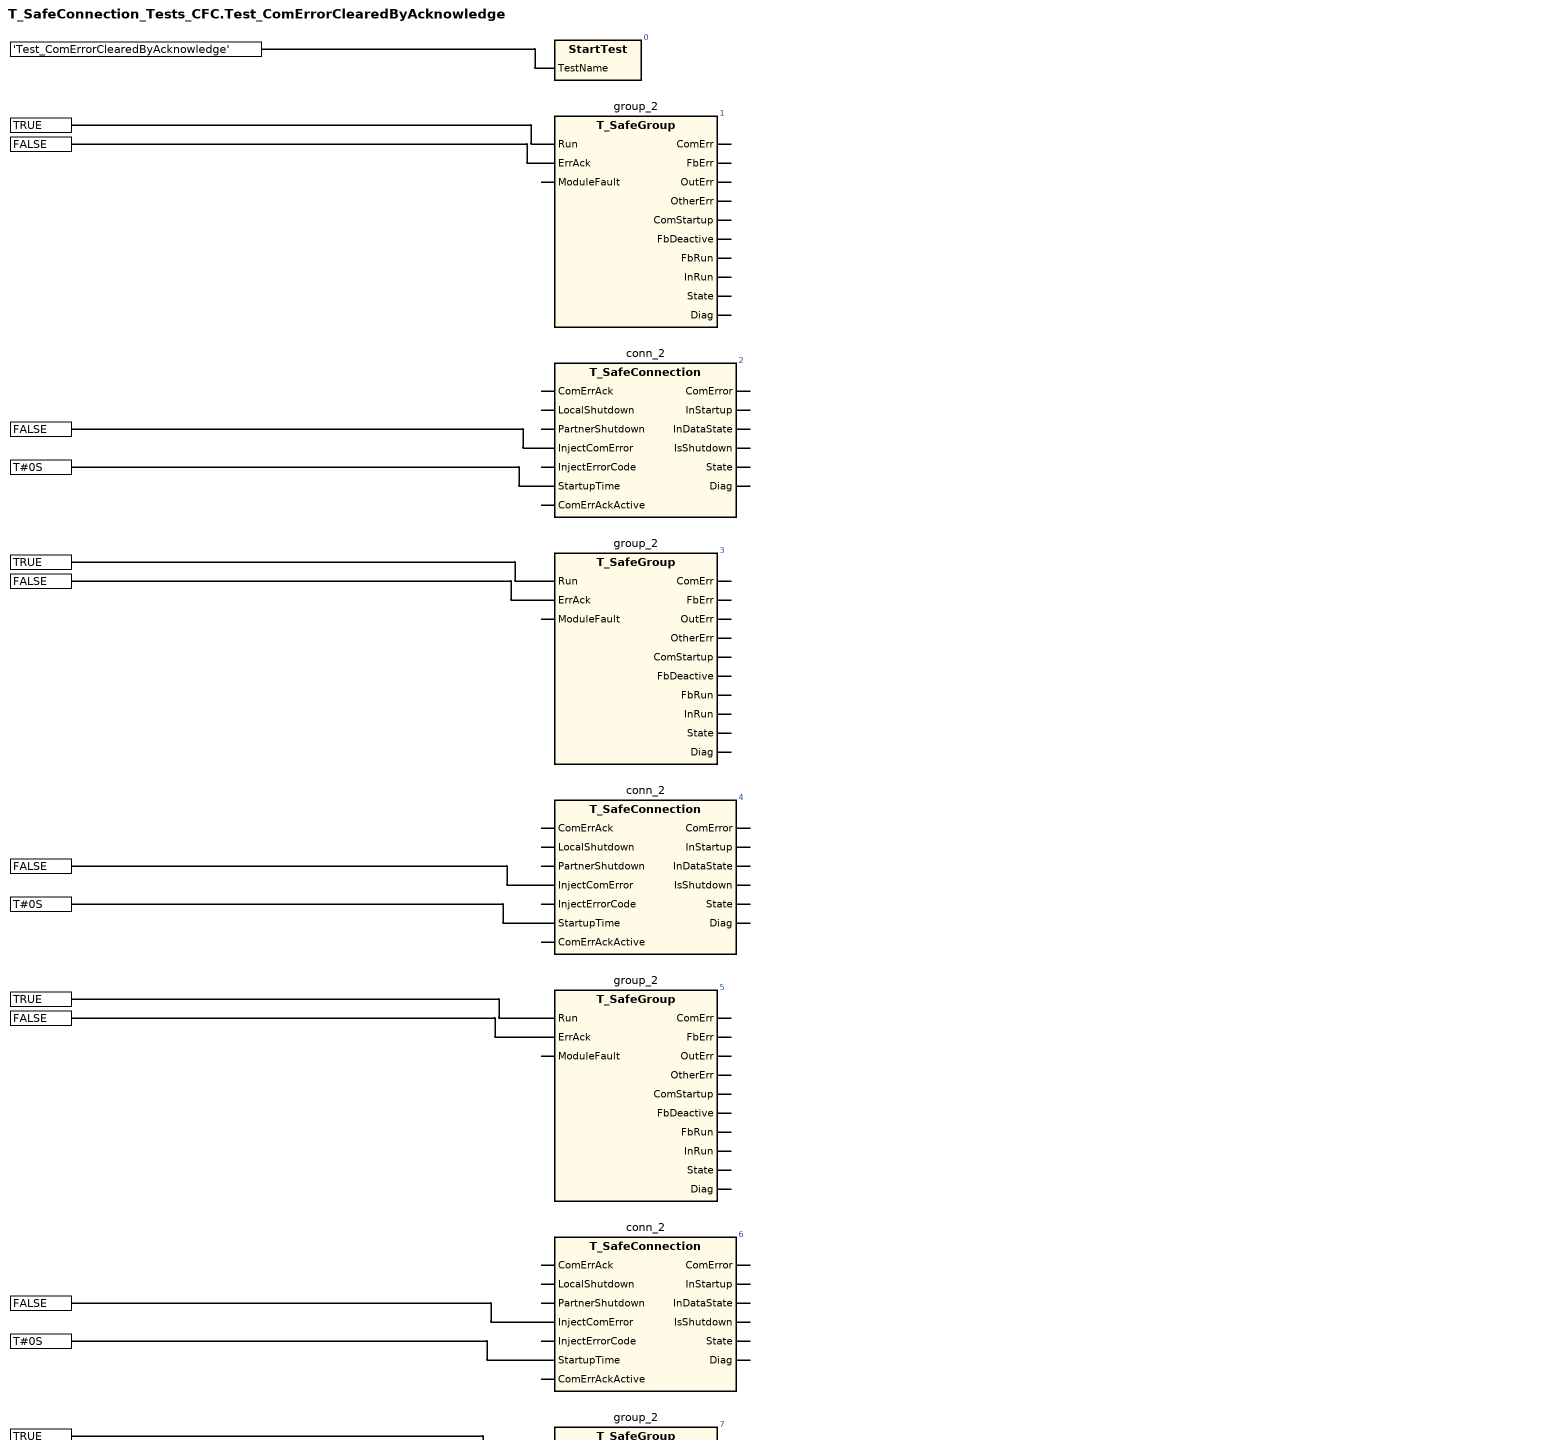
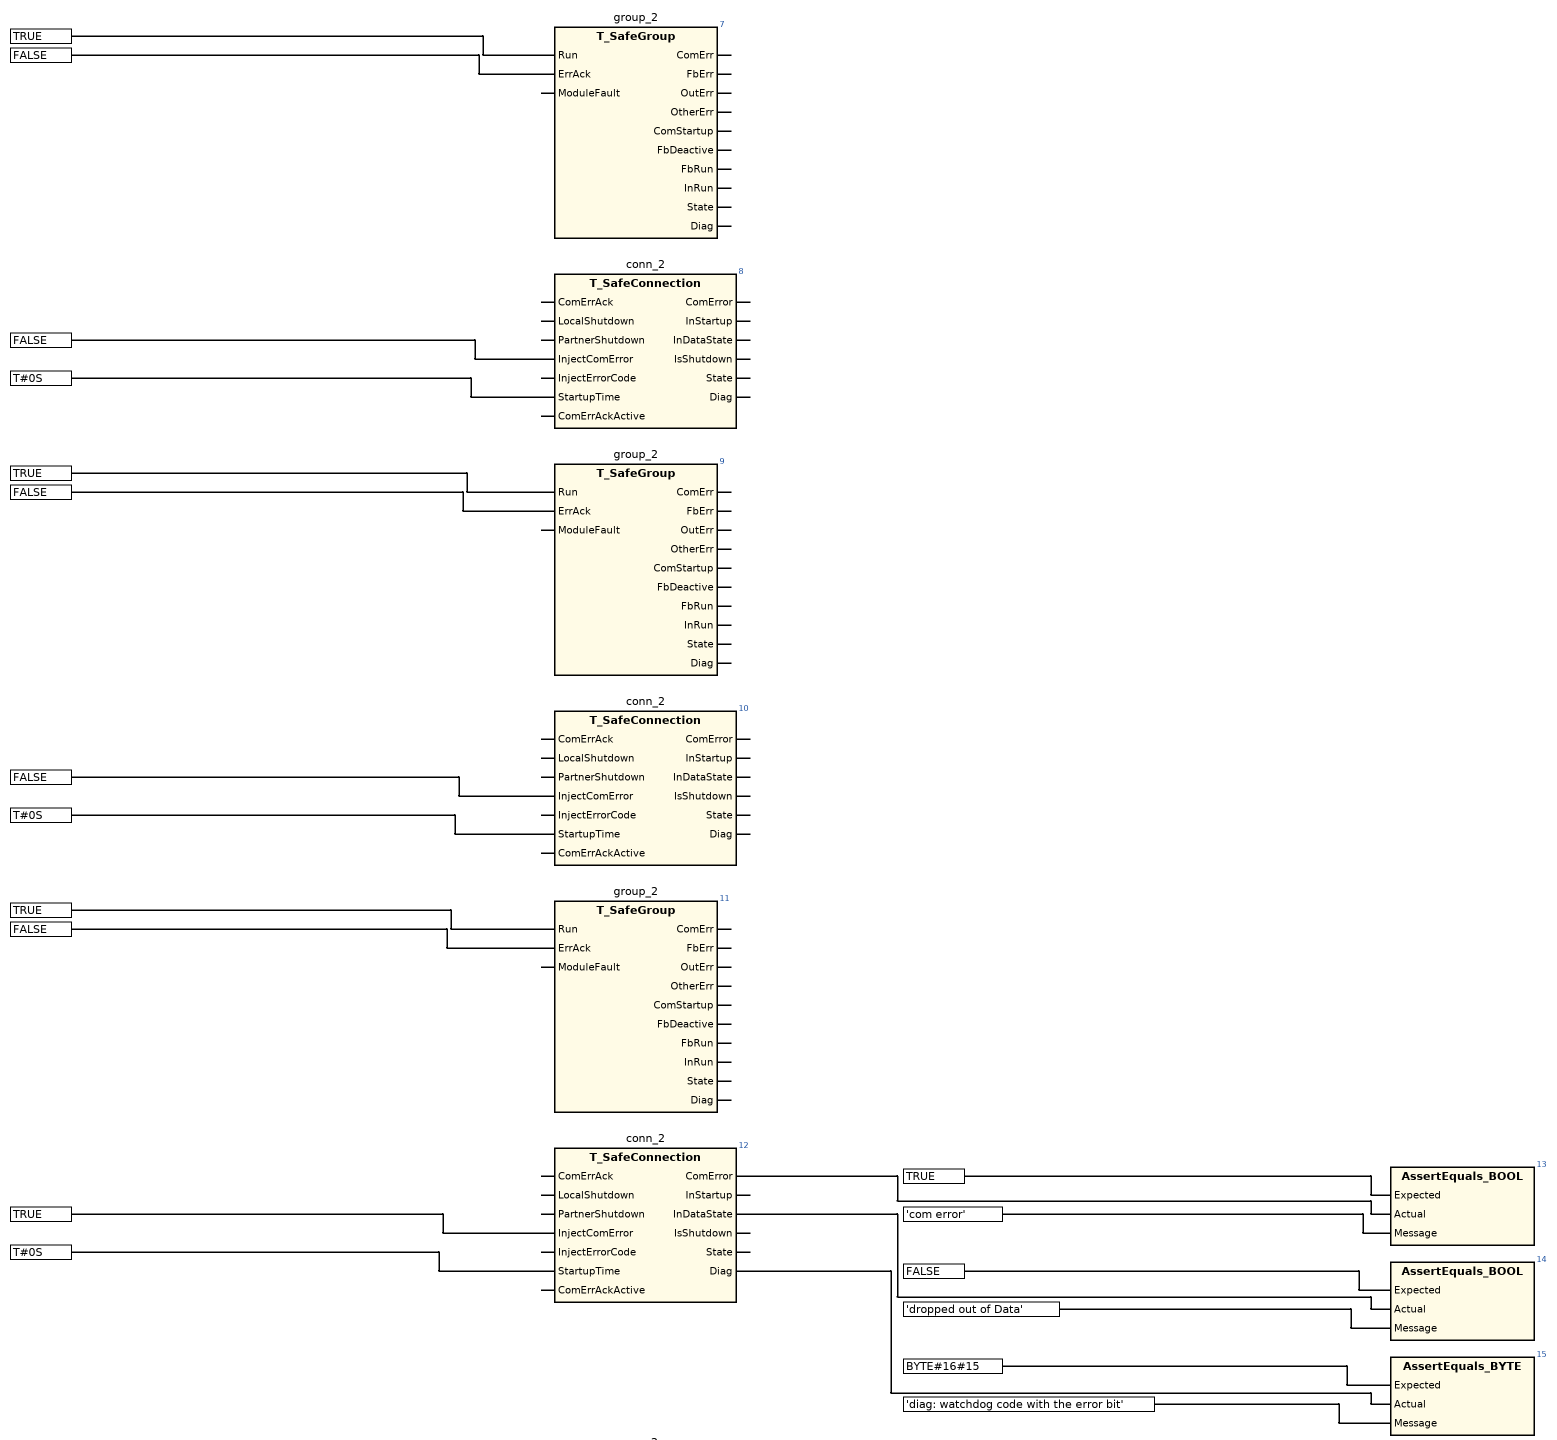
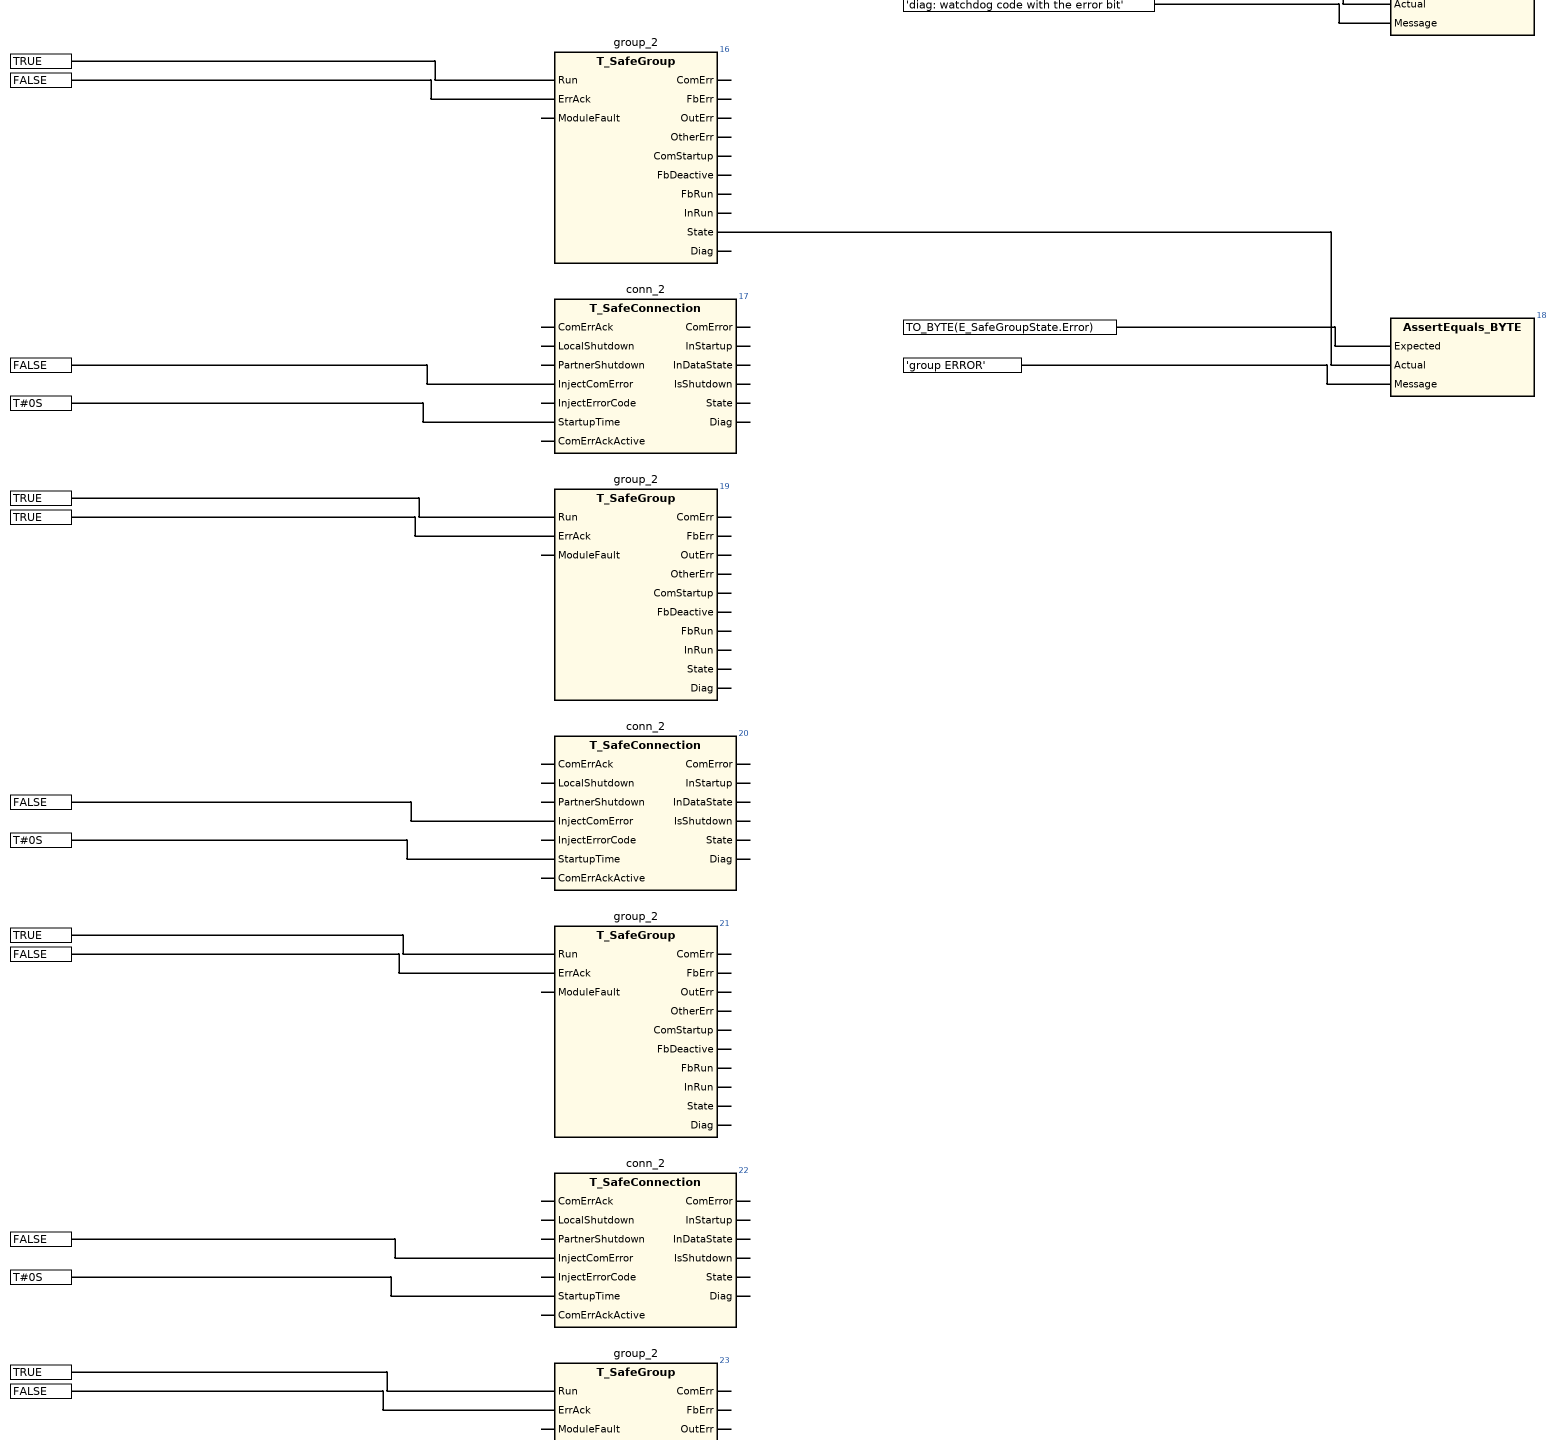
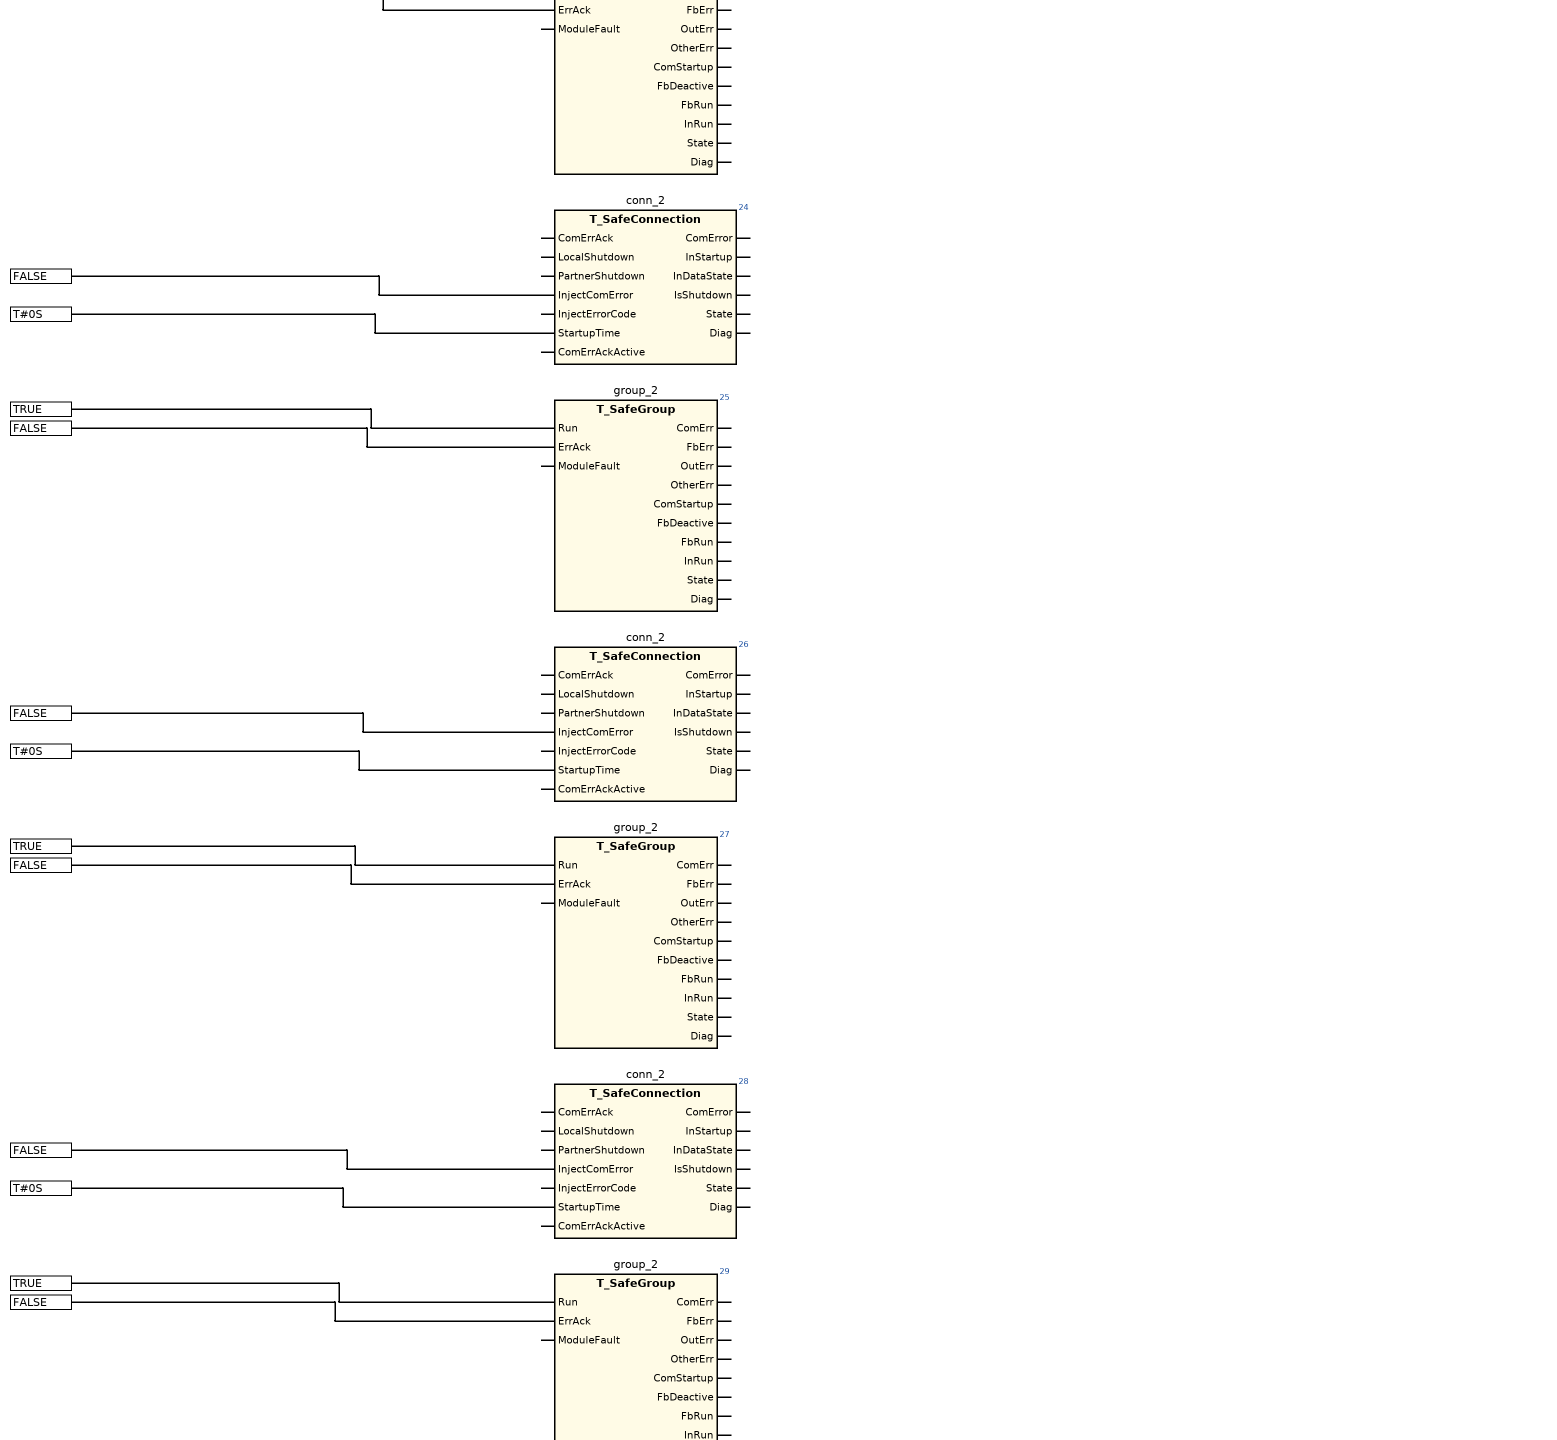
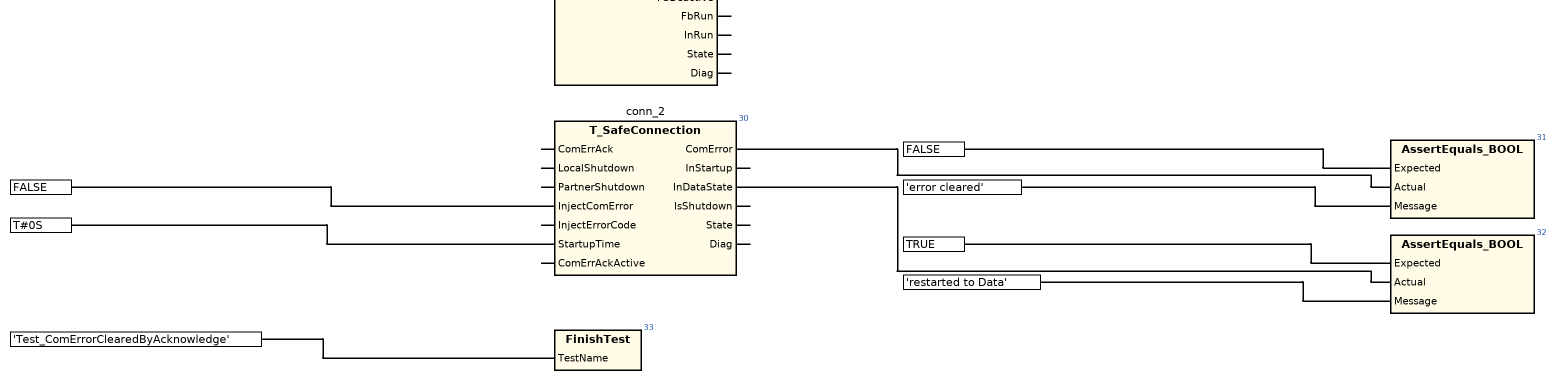
StartTest(TestName := 'Test_ComErrorClearedByAcknowledge');
group_2(Run := TRUE, ErrAck := FALSE); // T_SafeGroup
conn_2(InjectComError := FALSE, StartupTime := T#0S); // T_SafeConnection
group_2(Run := TRUE, ErrAck := FALSE); // T_SafeGroup
conn_2(InjectComError := FALSE, StartupTime := T#0S); // T_SafeConnection
group_2(Run := TRUE, ErrAck := FALSE); // T_SafeGroup
conn_2(InjectComError := FALSE, StartupTime := T#0S); // T_SafeConnection
group_2(Run := TRUE, ErrAck := FALSE); // T_SafeGroup
conn_2(InjectComError := FALSE, StartupTime := T#0S); // T_SafeConnection
group_2(Run := TRUE, ErrAck := FALSE); // T_SafeGroup
conn_2(InjectComError := FALSE, StartupTime := T#0S); // T_SafeConnection
group_2(Run := TRUE, ErrAck := FALSE); // T_SafeGroup
conn_2(InjectComError := TRUE, StartupTime := T#0S); // T_SafeConnection
AssertEquals_BOOL(Expected := TRUE, Actual := conn_2.ComError, Message := 'com error');
AssertEquals_BOOL(Expected := FALSE, Actual := conn_2.InDataState, Message := 'dropped out of Data');
AssertEquals_BYTE(Expected := BYTE#16#15, Actual := conn_2.Diag, Message := 'diag: watchdog code with the error bit');
group_2(Run := TRUE, ErrAck := FALSE); // T_SafeGroup
conn_2(InjectComError := FALSE, StartupTime := T#0S); // T_SafeConnection
AssertEquals_BYTE(Expected := TO_BYTE(E_SafeGroupState.Error), Actual := group_2.State, Message := 'group ERROR');
group_2(Run := TRUE, ErrAck := TRUE); // T_SafeGroup
conn_2(InjectComError := FALSE, StartupTime := T#0S); // T_SafeConnection
group_2(Run := TRUE, ErrAck := FALSE); // T_SafeGroup
conn_2(InjectComError := FALSE, StartupTime := T#0S); // T_SafeConnection
group_2(Run := TRUE, ErrAck := FALSE); // T_SafeGroup
conn_2(InjectComError := FALSE, StartupTime := T#0S); // T_SafeConnection
group_2(Run := TRUE, ErrAck := FALSE); // T_SafeGroup
conn_2(InjectComError := FALSE, StartupTime := T#0S); // T_SafeConnection
group_2(Run := TRUE, ErrAck := FALSE); // T_SafeGroup
conn_2(InjectComError := FALSE, StartupTime := T#0S); // T_SafeConnection
group_2(Run := TRUE, ErrAck := FALSE); // T_SafeGroup
conn_2(InjectComError := FALSE, StartupTime := T#0S); // T_SafeConnection
AssertEquals_BOOL(Expected := FALSE, Actual := conn_2.ComError, Message := 'error cleared');
AssertEquals_BOOL(Expected := TRUE, Actual := conn_2.InDataState, Message := 'restarted to Data');
FinishTest(TestName := 'Test_ComErrorClearedByAcknowledge');
END_METHOD

METHOD PRIVATE Test_StartsUpToDataWhenGroupRuns
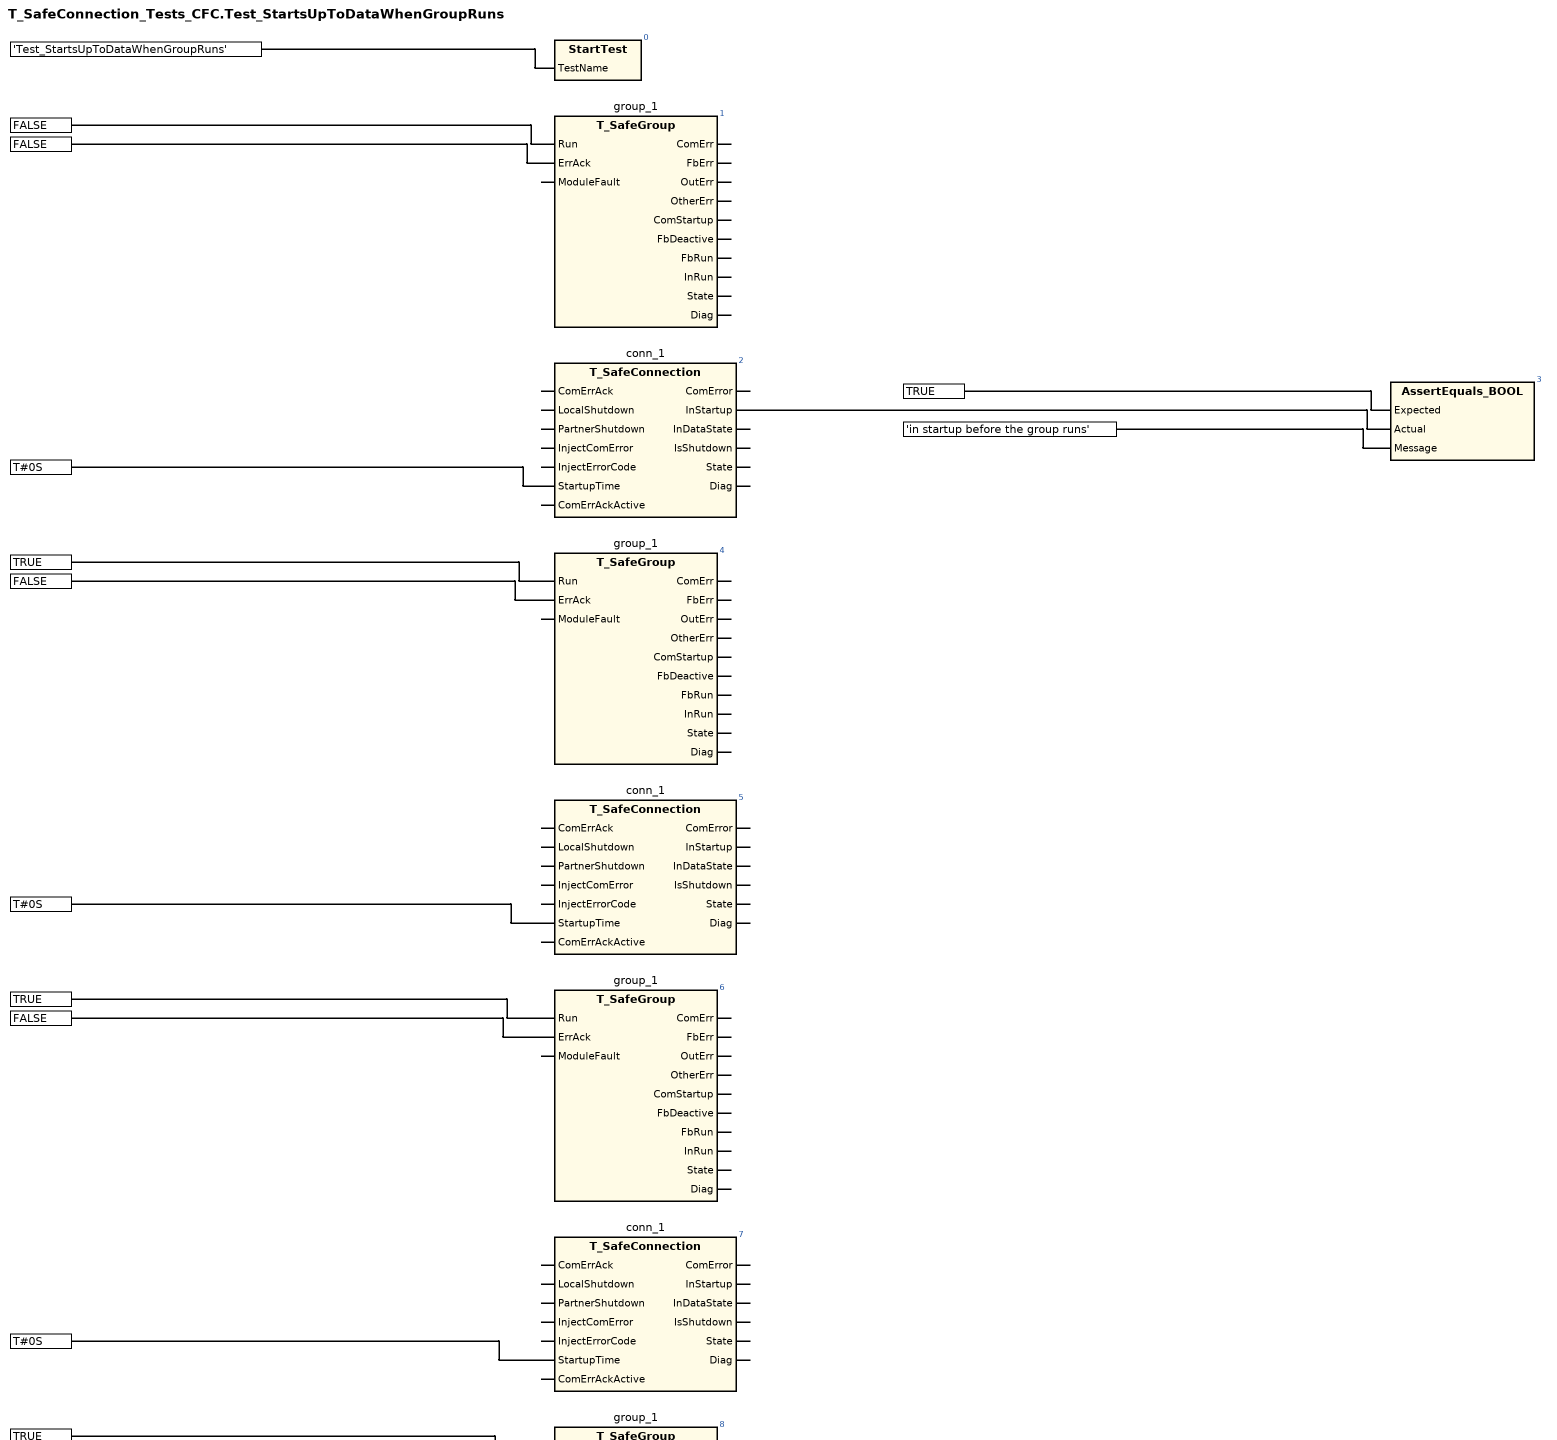
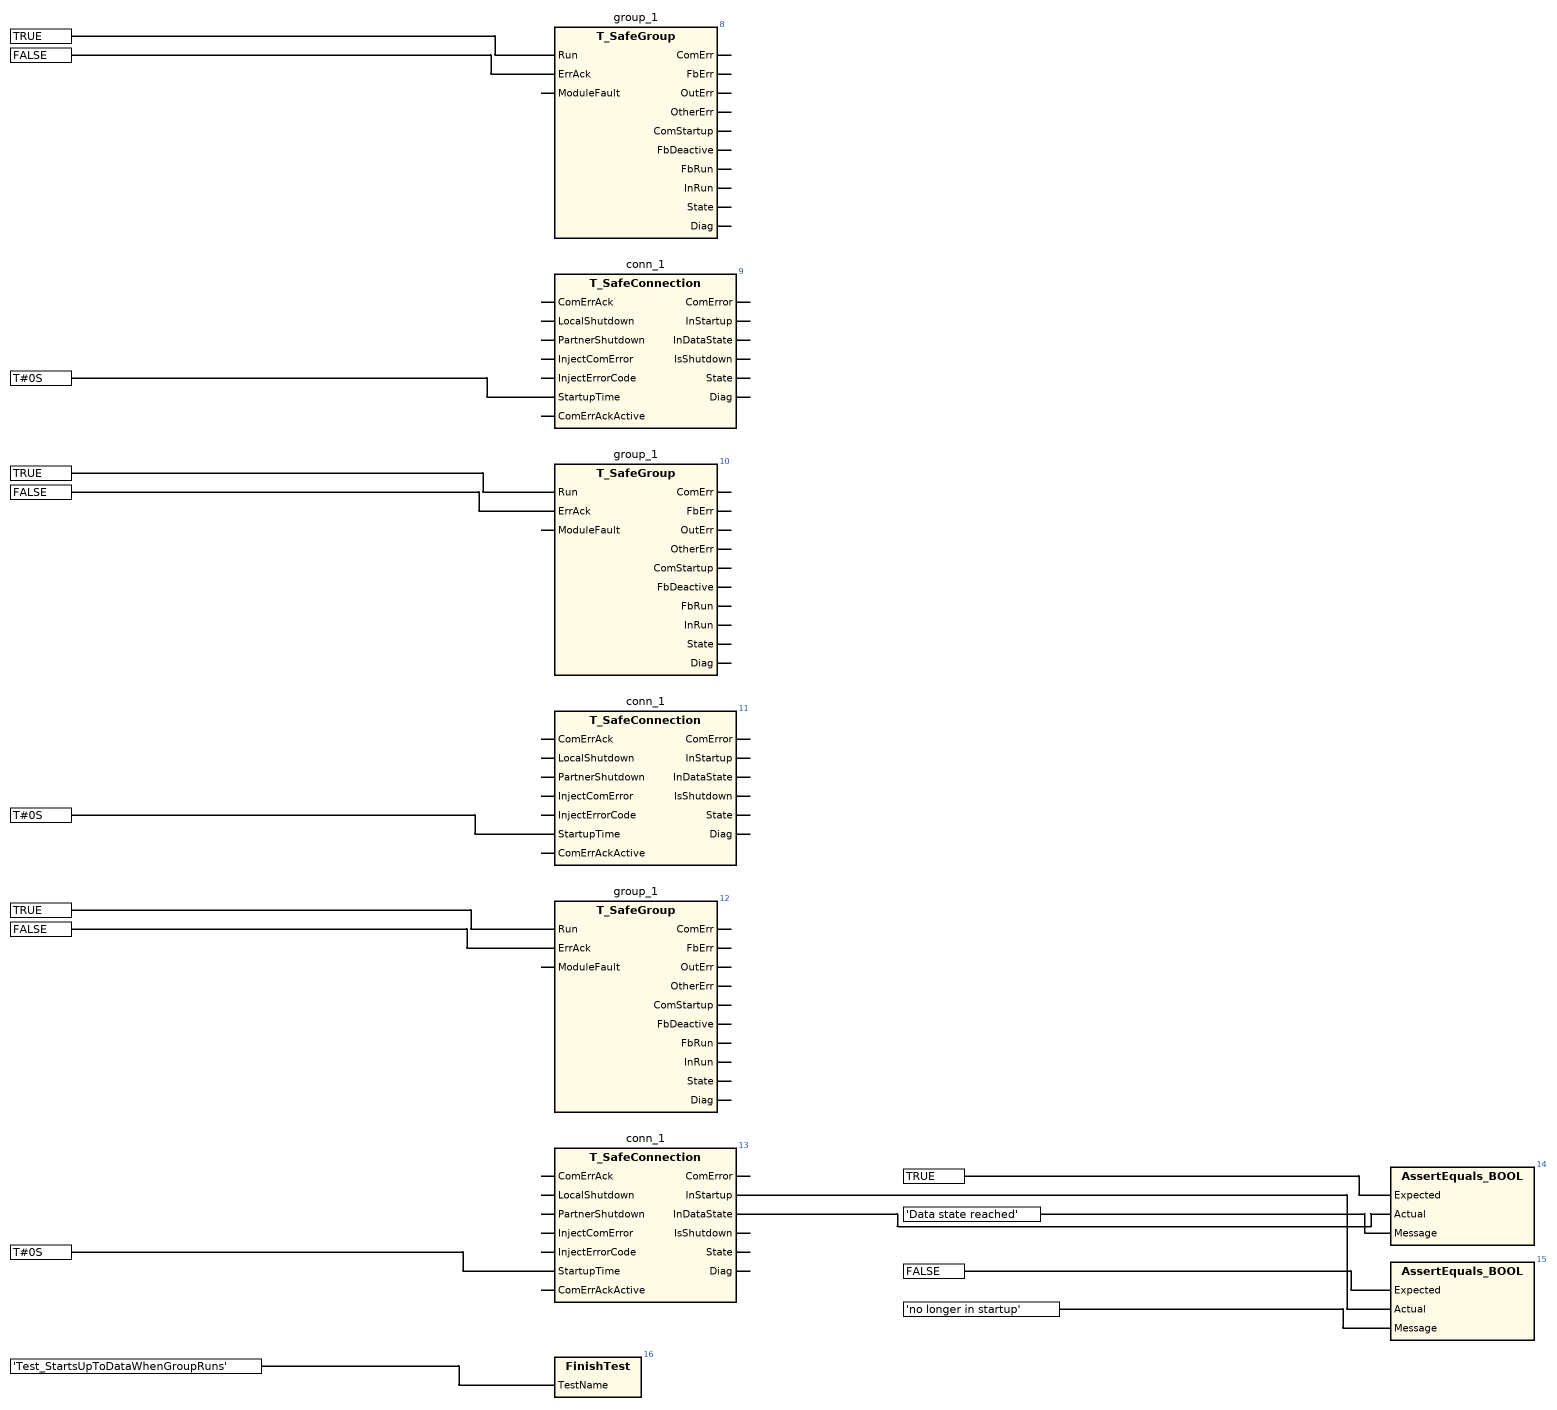
StartTest(TestName := 'Test_StartsUpToDataWhenGroupRuns');
group_1(Run := FALSE, ErrAck := FALSE); // T_SafeGroup
conn_1(StartupTime := T#0S); // T_SafeConnection
AssertEquals_BOOL(Expected := TRUE, Actual := conn_1.InStartup, Message := 'in startup before the group runs');
group_1(Run := TRUE, ErrAck := FALSE); // T_SafeGroup
conn_1(StartupTime := T#0S); // T_SafeConnection
group_1(Run := TRUE, ErrAck := FALSE); // T_SafeGroup
conn_1(StartupTime := T#0S); // T_SafeConnection
group_1(Run := TRUE, ErrAck := FALSE); // T_SafeGroup
conn_1(StartupTime := T#0S); // T_SafeConnection
group_1(Run := TRUE, ErrAck := FALSE); // T_SafeGroup
conn_1(StartupTime := T#0S); // T_SafeConnection
group_1(Run := TRUE, ErrAck := FALSE); // T_SafeGroup
conn_1(StartupTime := T#0S); // T_SafeConnection
AssertEquals_BOOL(Expected := TRUE, Actual := conn_1.InDataState, Message := 'Data state reached');
AssertEquals_BOOL(Expected := FALSE, Actual := conn_1.InStartup, Message := 'no longer in startup');
FinishTest(TestName := 'Test_StartsUpToDataWhenGroupRuns');
END_METHOD

END_FUNCTION_BLOCK

// Tests/T_SafeConnShutdown_Tests_CFC
    // CFC twin of T_SafeConnShutdown_Tests: the same tests drawn as CFC diagrams, the way a TwinSAFE project is authored.
    FUNCTION_BLOCK T_SafeConnShutdown_Tests_CFC EXTENDS T_SafeCfcTestSuite
    VAR
    // Test_DeactivateShutsDownConnection
    group_1 : T_SafeGroup;
    conn_1 : T_SafeConnection(group := group_1);
    fb_1 : T_SafeConnShutdown(group := group_1, connection := conn_1);
END_VAR

Test_DeactivateShutsDownConnection();

METHOD PRIVATE Test_DeactivateShutsDownConnection
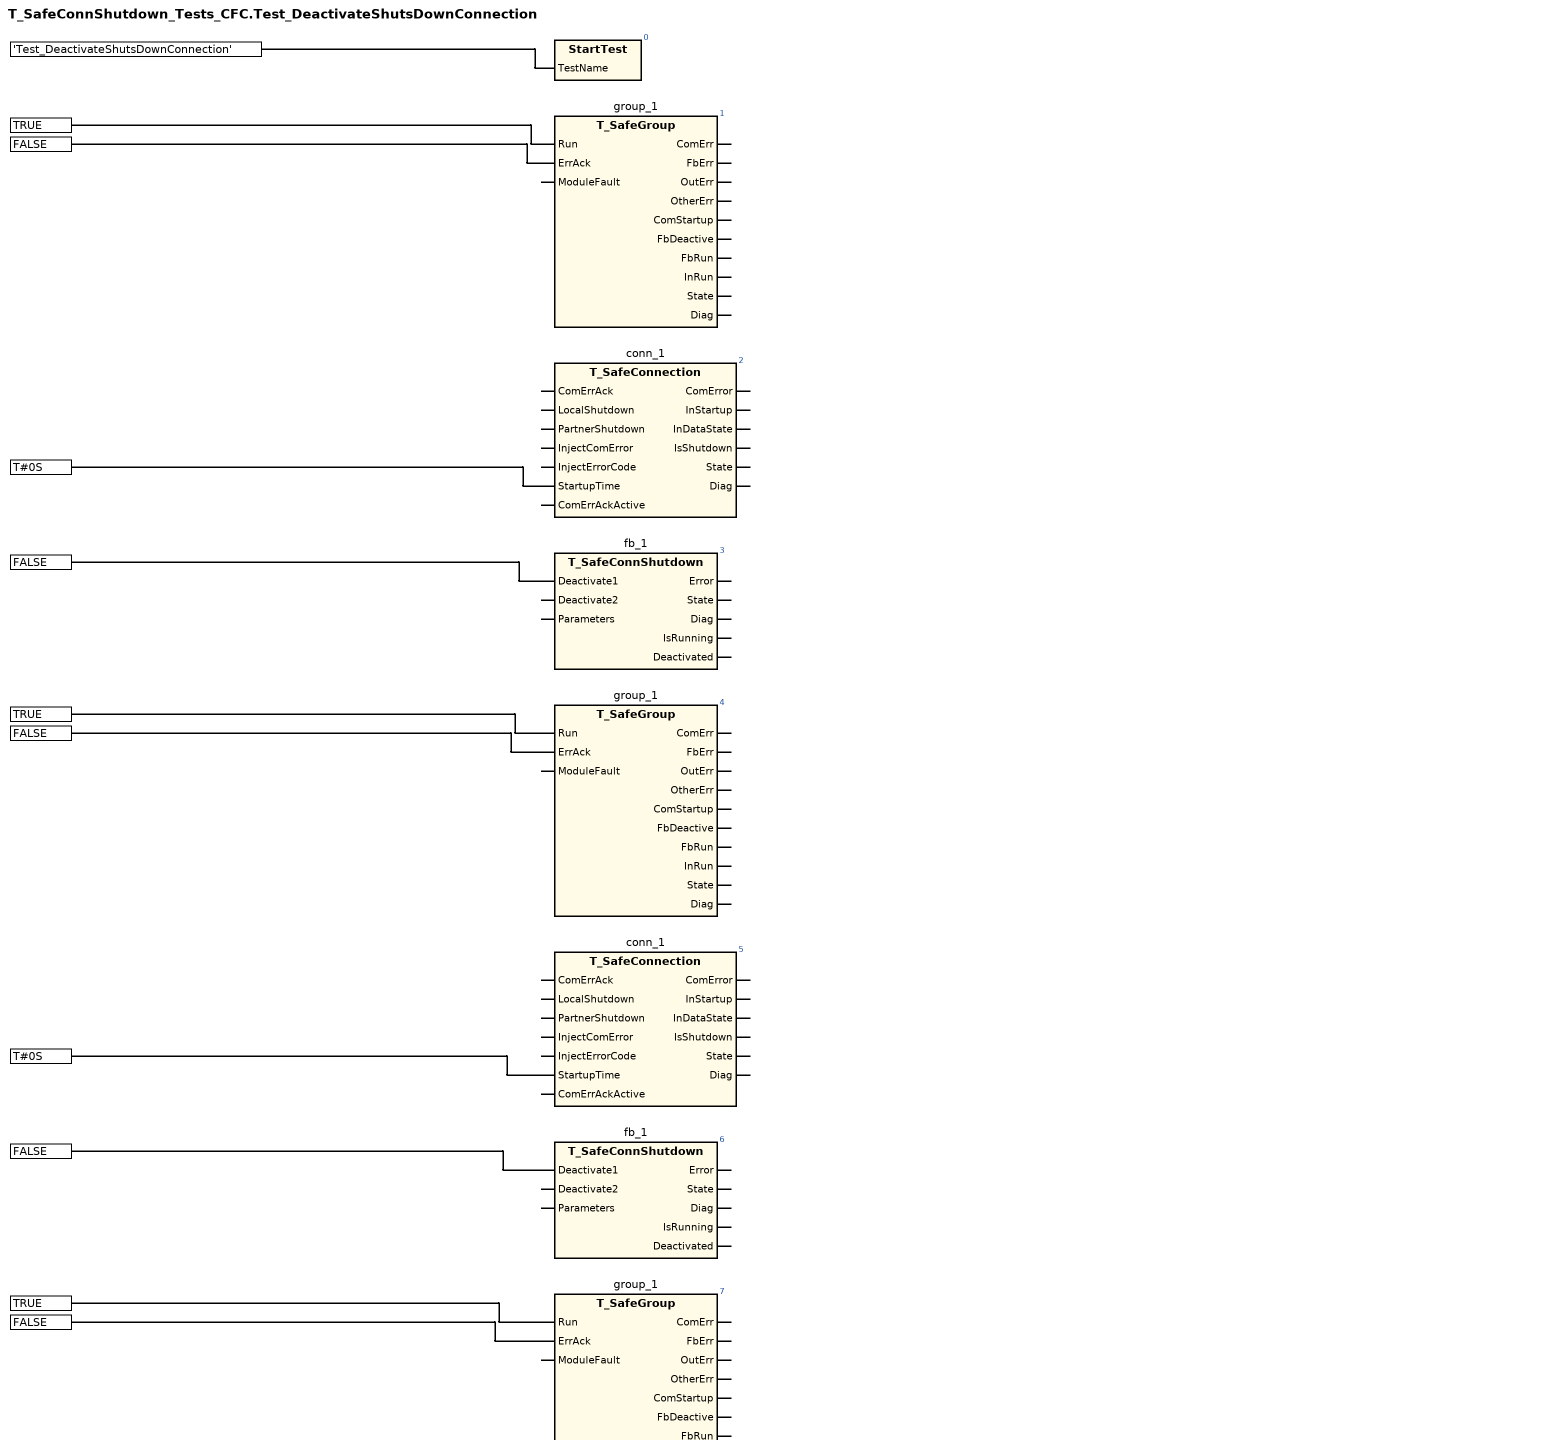
